  def gripper_to_mm(value_gripper, gripper_socket):
      closed_norm = get_closed_norm(gripper_socket)
      open_norm = get_open_norm(gripper_socket)
      closed_mm = get_closed_mm(gripper_socket)
      open_mm = get_open_mm(gripper_socket)

      value_norm = (value_gripper / 255) * 100

      slope = (closed_mm - open_mm) / (closed_norm - open_norm)
      value_mm = slope * (value_norm - closed_norm) + closed_mm

      if (value_mm > open_mm):
          value_mm_limited = open_mm
      elif (value_mm < closed_mm):
          value_mm_limited = closed_mm
      else:
          value_mm_limited = value_mm
      end

      return value_mm_limited
  end

  def mm_to_gripper(value_mm, gripper_socket):
      closed_norm = get_closed_norm(gripper_socket)
      open_norm = get_open_norm(gripper_socket)
      closed_mm = get_closed_mm(gripper_socket)
      open_mm = get_open_mm(gripper_socket)

      slope = (closed_norm - open_norm) / (closed_mm - open_mm)
      value_norm = (value_mm - closed_mm) * slope + closed_norm

      value_gripper = value_norm * 255 / 100

      if (value_gripper > 255):
          value_gripper_limited = 255
      elif (value_gripper < 0):
          value_gripper_limited = 0
      else:
          value_gripper_limited = round_value(value_gripper)
      end

      return value_gripper_limited
  end

  def round_value(value):
      value_mod = value % 1

      if(value_mod < 0.5):
          return floor(value)
      else:
          return ceil(value)
      end
  end

  def round_value_2_dec(value):
      value_x_100 = value * 100
      value_x_100_rounded = round_value(value_x_100)
      return value_x_100_rounded / 100
  end

  def clear_socket_buffer(gripper_socket="1", read_timeout = 0.1):
      rq_comm_clear_socket_buffer_enabled[rq_socket_to_index(gripper_socket)] = True
  end

  def rq_gripper_id_to_ascii(gripper_id):
      if(gripper_id == "1"):
          return 57
      elif(gripper_id == "2"):
          return 50
      elif(gripper_id == "3"):
          return 51
      elif(gripper_id == "4"):
          return 52
      end
  end

      def scale(value, rawRange, scaledRange):
          def computeSlope(inputRange, outputRange):
              outputRangeDelta = outputRange[1] - outputRange[0]
              inputRangeDelta = inputRange[1] - inputRange[0]

              if (inputRangeDelta == 0):
                  return 0
              else:
                  return outputRangeDelta / inputRangeDelta
              end
          end

          def computeIntercept(slope, inputRange, outputRange):
              return outputRange[0] - (slope * inputRange[0])
          end

          def clipScaledValue(outputScaledValue, outputRange):
              if (outputRange[0] < outputRange[1]):
                  return clipWhenLowerLimitIsLessThanHigher(outputScaledValue, outputRange)
              else:
                  return clipWhenLowerLimitIsGreaterThanHigherLimit(outputScaledValue, outputRange)
              end
          end

          def clipWhenLowerLimitIsGreaterThanHigherLimit(outputScaledValue, outputRange):
              if (outputScaledValue < outputRange[1]):
                  return outputRange[1]
              elif (outputScaledValue > outputRange[0]):
                  return outputRange[0]
              else:
                  return outputScaledValue
              end
          end

          def clipWhenLowerLimitIsLessThanHigher(outputScaledValue, outputRange):
              if (outputScaledValue < outputRange[0]):
                  return outputRange[0]
              elif (outputScaledValue > outputRange[1]):
                  return outputRange[1]
              else:
                  return outputScaledValue
              end
          end

          slope = computeSlope(rawRange, scaledRange)
          intercept = computeIntercept(slope, rawRange, scaledRange)
          scaledValue = slope * value + intercept
          return clipScaledValue(scaledValue, scaledRange)
      end

      def limit(value, range):
          return scale(value, range, range)
      end


  rq_init_comm_if_connected(9, "1")
  rq_init_comm_if_connected(2, "2")
  rq_init_comm_if_connected(3, "3")
  rq_init_comm_if_connected(4, "4")
  rq_print_connected_grippers()
  rq_gripper_communication_thread = run rq_gripper_communication()
  set_closed_norm(97.6470588235294, "1")
  set_open_norm(1.1764705882352942, "1")
  set_closed_mm(0.0, "1")
  set_open_mm(53.0, "1")
  set_closed_norm(100.0, "2")
  set_open_norm(0.0, "2")
  set_closed_mm(0.0, "2")
  set_open_mm(50.0, "2")
  set_closed_norm(100.0, "3")
  set_open_norm(0.0, "3")
  set_closed_mm(0.0, "3")
  set_open_mm(50.0, "3")
  set_closed_norm(100.0, "4")
  set_open_norm(0.0, "4")
  set_closed_mm(0.0, "4")
  set_open_mm(50.0, "4")
  rq_current_limit_enabled = False
  while(not rq_gripper_communication_thread_started):
      sleep(0.008)
  end
  # end: URCap Installation Node
  step_count_af30497c_f8d6_4abb_9ab3_badfcb3aff49 = 0.0
  thread Step_Counter_Thread_6e0f90e9_d7f0_45c2_bba1_3f0a34dad08c():
    while (True):
      step_count_af30497c_f8d6_4abb_9ab3_badfcb3aff49 = step_count_af30497c_f8d6_4abb_9ab3_badfcb3aff49 + 1.0
      sync()
    end
  end
  run Step_Counter_Thread_6e0f90e9_d7f0_45c2_bba1_3f0a34dad08c()
  global AMR_Position=struct(position_identifier=0, x1=0, x2=0, y1=0, y2=0, theta1=0, theta2=0)
  global CAM_Pose=p[0,0,0,0,0,0]
  global CAM_Relation=""
  global CMD_Abort=  False
  global CMD_Clear=  False
  global CMD_Reset=  False
  global CMD_Start=  False
  global CMD_Suspend=  False
  global CMD_Unhold=  False
  global CMD_Unsuspend=  False
  global CNT_Rack_Output=0
  global FNC_Freedrive=  False
  global PRC_TubCounter=0
  global STP=0
  global easyPickCount_4=0
  global easyPickCount_7=0
  global easyPickNoObj_4=0
  global easyPickNoObj_7=0
  global easyPickParts_4=0
  global easyPickParts_7=0
  global TMR_Barcode=0
  global Container_mid_1_p=p[-.379239199143, -.127191311915, .299999999998, .000000000046, -.000000000021, -1.247199999994]
  global Container_mid_1_q=[-2.477408934449926, -1.2969853503591224, -1.875639182904262, -1.539621866126728, 1.5731943360401213, -2.8009955944022717]
  global trigger_otw_p=p[-.364831738276, -.163967193938, .343299997821, .000000000046, -.000000000020, -1.148401333327]
  global trigger_otw_q=[-2.378283213085033, -1.2994862387706814, -1.7634300687554951, -1.6493302004167063, 1.573123683454141, -2.8011223671816943]
  global Waypoint_54_p=p[.008800512419, -.547926542621, .402696567415, -.589884378425, -.007228654778, -.061268144704]
  global Waypoint_54_q=[-1.2044575850116175, -1.3416667741588135, -1.8272563219070435, -0.9884541195682068, 1.3621035814285278, -2.7712565104113978]
  global Waypoint_77_p=p[-.178371829612, -.433927395311, .368082383916, -.086593488055, .704679941724, -.007869906074]
  global Waypoint_77_q=[-1.265390698109762, -1.3355963987163086, -1.7944865226745605, -1.7402602634825648, 0.8780410885810852, -2.7713127771960657]
  global Waypoint_83_p=p[.008800512419, -.547926542621, .402696567415, -.589884378425, -.007228654778, -.061268144704]
  global Waypoint_83_q=[-1.2044575850116175, -1.3416667741588135, -1.8272563219070435, -0.9884541195682068, 1.3621035814285278, -2.7712565104113978]
  global Waypoint_84_p=p[-.178371829612, -.433927395311, .368082383916, -.086593488055, .704679941724, -.007869906074]
  global Waypoint_84_q=[-1.265390698109762, -1.3355963987163086, -1.7944865226745605, -1.7402602634825648, 0.8780410885810852, -2.7713127771960657]
  global Vial_above_1_p=p[.017105793010, -.652093028359, .184920586844, .000000000272, .000000000270, 1.564063451276]
  global Vial_above_1_q=[-1.3375440709712851, -1.9618096977868804, -1.4665759083780685, -1.2837941559171444, 1.5732503672317195, -4.47276330421513]
  global Vial_pick_poi_1_p=p[.017105792852, -.648922724010, .093307568731, .000000000271, .000000000270, 1.564063451276]
  global Vial_pick_poi_1_q=[-1.3366329456391917, -2.0375277831965413, -1.6071432798879028, -1.0675084332049813, 1.57309887265915, -4.471135348858068]
  global Waypoint_86_p=p[.019227646885, -.648669633640, .184920586950, .000000000000, .000000000000, .024063451426]
  global Waypoint_86_q=[-1.3331129109407733, -1.9540750545686123, -1.4775914902901128, -1.280581784992414, 1.5733500744865856, -2.928303704452631]
  global Waypoint_87_p=p[-.032361834699, -.348336136197, .391475576335, -.000008499254, .000014589902, -.004651426820]
  global Waypoint_87_q=[-1.2709335019096129, -1.1914598663441005, -1.708995335060501, -1.8117888533498316, 1.5729683532263925, -2.8379347397710237]
  global Vial_3FG_plac_1_p=p[-.031858676359, -.349402499566, .145301120695, .000000000000, .000000000000, .000000000000]
  global Vial_3FG_plac_1_q=[-1.2723975525801707, -1.252376585823825, -2.3128114007049496, -1.1470592278900167, 1.5730548099411423, -2.8414815174610535]
  global Waypoint_88_p=p[-.032361834699, -.348336136197, .391475576335, -.000008499254, .000014589902, -.004651426820]
  global Waypoint_88_q=[-1.2709335019096129, -1.1914598663441005, -1.708995335060501, -1.8117888533498316, 1.5729683532263925, -2.8379347397710237]
  global cap_dump_1_p=p[-.139168676487, -.420163541420, .146096395183, .000000000000, .000000000000, .000000000000]
  global cap_dump_1_q=[-1.584588644510994, -1.5093464179777323, -2.1118449369620347, -1.091059703602438, 1.5728943834877336, -3.154014906686923]
  global Waypoint_89_p=p[-.032361834699, -.348336136197, .391475576335, -.000008499254, .000014589902, -.004651426820]
  global Waypoint_89_q=[-1.2709335019096129, -1.1914598663441005, -1.708995335060501, -1.8117888533498316, 1.5729683532263925, -2.8379347397710237]
  global Vial_3FG_plac_2_p=p[-.031858676359, -.349402499566, .145301120695, .000000000000, .000000000000, .000000000000]
  global Vial_3FG_plac_2_q=[-1.2723975525801707, -1.252376585823825, -2.3128114007049496, -1.1470592278900167, 1.5730548099411423, -2.8414815174610535]
  global Waypoint_90_p=p[-.032361834699, -.348336136197, .391475576335, -.000008499254, .000014589902, -.004651426820]
  global Waypoint_90_q=[-1.2709335019096129, -1.1914598663441005, -1.708995335060501, -1.8117888533498316, 1.5729683532263925, -2.8379347397710237]
  global cap_dump_2_p=p[-.139168676487, -.420163541420, .146096395183, .000000000000, .000000000000, .000000000000]
  global cap_dump_2_q=[-1.584588644510994, -1.5093464179777323, -2.1118449369620347, -1.091059703602438, 1.5728943834877336, -3.154014906686923]
  global Waypoint_91_p=p[-.032361834699, -.348336136197, .391475576335, -.000008499254, .000014589902, -.004651426820]
  global Waypoint_91_q=[-1.2709335019096129, -1.1914598663441005, -1.708995335060501, -1.8117888533498316, 1.5729683532263925, -2.8379347397710237]
  global Vial_liq_abov_1_p=p[-.025303660977, -.338758622354, .426628485936, -1.315858642253, .800043520260, -.928295855026]
  global Vial_liq_abov_1_q=[-0.3789628187762659, -1.5149522957256814, -2.263045310974121, 0.7870649534412841, -0.750984017048971, -3.2237566153155726]
  global Vial_liq_pick_3_p=p[-.002660428945, -.335984893034, .159389832934, -1.150456778400, .673175527684, -1.010612657503]
  global Vial_liq_pick_3_q=[-0.3660772482501429, -1.4503649038127442, -2.4056053161621094, -1.994692941705221, 0.8039668202400208, -0.2508929411517542]
  global Vial_liq_pick_4_p=p[-.041402486291, -.356791603314, .125395323246, -1.143483969075, .651070210027, -.878721885453]
  global Vial_liq_pick_4_q=[-0.4426233705502476, -1.437252121513727, -2.551930962114307, -1.776528229806984, 0.6562026234073748, -0.43018811960029524]
  global Vial_liq_abov_2_p=p[-.025303660977, -.338758622354, .426628485936, -1.315858642253, .800043520260, -.928295855026]
  global Vial_liq_abov_2_q=[-0.3789628187762659, -1.5149522957256814, -2.263045310974121, 0.7870649534412841, -0.750984017048971, -3.2237566153155726]
  global Liquid_midway_1_p=p[.057575295009, -.583081747994, .306414980749, -1.351675548728, .120935756539, -.096908606303]
  global Liquid_midway_1_q=[-0.895174805318014, -1.7035466633238734, -2.380953073501587, 0.631549521083496, 0.7706599235534668, -2.9455552736865442]
  global shake_3_p=p[.057574880217, -.583085370269, .306422893466, -1.360996190983, -.155555042453, -.438136255921]
  global shake_3_q=[-0.8951800505267542, -1.7035466633238734, -2.380937099456787, 0.6315542894550782, 0.7706599235534669, -2.5394540616517496]
  global shake_4_p=p[.057581636113, -.583090570002, .306439684073, -1.308767904323, .368530312677, .214926493520]
  global shake_4_q=[-0.8951714674579065, -1.7035395107665003, -2.380906343460083, 0.6315504747578125, 0.7706480026245118, -3.3161255787892268]
  global drop_above_3_p=p[.268235025993, -.467784390499, .226219872376, -1.027832627524, -.430841408251, 1.004603115937]
  global drop_above_3_q=[-0.935645882283346, -1.6663371525206507, -2.4252893924713135, 0.41966931402172847, 1.8470635414123535, -3.4600217978106897]
  global drop_above_4_p=p[.219042229014, -.470775657081, .133754190740, -.313004595901, -.344395319364, 1.500564994056]
  global drop_above_4_q=[-1.0601594887284795, -1.70046459045642, -2.0799996233759863, -0.7243227230676759, 1.9429634314685202, -4.115129153870795]
  global liq_tran_3_p=p[.213067510942, -.469567035397, .100231043184, .251862243732, .217902579404, 1.592812335393]
  global liq_tran_3_q=[-0.7789645168037476, -1.822364827406652, -1.8643518410805573, -1.252158963840138, 1.3768134449520435, -3.9328333233290254]
  global drop_above_5_p=p[.219042229014, -.470775657081, .133754190740, -.313004595901, -.344395319364, 1.500564994056]
  global drop_above_5_q=[-1.0601594887284795, -1.70046459045642, -2.0799996233759863, -0.7243227230676759, 1.9429634314685202, -4.115129153870795]
  global Waypoint_92_p=p[.187119460405, -.493959476151, .133754190608, -.313004596540, -.344395317757, 1.500564993991]
  global Waypoint_92_q=[-1.1418328121400876, -1.7310553375189475, -2.033634768766424, -0.772026910513711, 1.958578934631971, -4.201588449364511]
  global liq_tran_4_p=p[.195957706507, -.493022614126, .100231042689, .160718757180, .109807038912, 1.525321508623]
  global liq_tran_4_q=[-0.881740380645474, -1.8244526267589851, -1.865100964490387, -1.1608866323693583, 1.4631433601076713, -3.973915130363038]
  global drop_above_6_p=p[.219042229014, -.470775657081, .133754190740, -.313004595901, -.344395319364, 1.500564994056]
  global drop_above_6_q=[-1.0601594887284795, -1.70046459045642, -2.0799996233759863, -0.7243227230676759, 1.9429634314685202, -4.115129153870795]
  global drop_above_7_p=p[.268235025993, -.467784390499, .226219872376, -1.027832627524, -.430841408251, 1.004603115937]
  global drop_above_7_q=[-0.935645882283346, -1.6663371525206507, -2.4252893924713135, 0.41966931402172847, 1.8470635414123535, -3.4600217978106897]
  global Liquid_midway_2_p=p[.057575295009, -.583081747994, .306414980749, -1.351675548728, .120935756539, -.096908606303]
  global Liquid_midway_2_q=[-0.895174805318014, -1.7035466633238734, -2.380953073501587, 0.631549521083496, 0.7706599235534668, -2.9455552736865442]
  global Vial_drop_abo_1_p=p[.000324902251, -.648569523142, .221894115667, -.873462921366, 1.165852672573, -1.482720593185]
  global Vial_drop_abo_1_q=[-1.0576906334721352, -2.393016994184633, -0.9236232851859159, -2.5729213042279273, 0.7903331288549689, -0.33286325848155585]
  global Vial_liq_drop_1_p=p[.001020867953, -.647659915585, .092915870838, -.834762611599, 1.081942994823, -1.540647900176]
  global Vial_liq_drop_1_q=[-1.0631954168193474, -2.4447642951220825, -1.128811017825127, -2.1983115491972294, 0.8130148661460634, -0.38984988696911316]
  global Vial_drop_abo_2_p=p[.000324902251, -.648569523142, .221894115667, -.873462921366, 1.165852672573, -1.482720593185]
  global Vial_drop_abo_2_q=[-1.0576906334721352, -2.393016994184633, -0.9236232851859159, -2.5729213042279273, 0.7903331288549689, -0.33286325848155585]
  global Spatula_otw_p=p[-.038472058237, -.263141484147, .425351216717, -.000441582511, -.000128175490, 3.034387645854]
  global Spatula_otw_q=[-1.1888947506684495, -1.0083288774886814, -1.7052227056065874, -1.9984805067363443, 1.5730180972985317, 0.48793409320312264]
  global pick_spat_L_abv_p=p[.239059466375, -.067212518441, .280720723617, .000017217488, -.000484427718, 3.106837214660]
  global pick_spat_L_abv_q=[0.292765616142962, -0.8565557553273315, -2.140199892763044, -1.715349495646084, 1.573623142106424, 1.8984976776985687]
  global spat_L_pick_p=p[.242468789885, -.067301915011, .193171208067, .000017217488, -.000484427718, 3.106837214657]
  global spat_L_pick_q=[0.2867414378807389, -0.8600077002089179, -2.3629148016312627, -1.4891831672860159, 1.5737695566221115, 1.8933890858591198]
  global spat_L_lift_p=p[.245402002494, -.067432373551, .289049296496, .000017217490, -.000484427724, 3.106837214657]
  global spat_L_lift_q=[0.2834351187564135, -0.8798320076811592, -2.1119436738532986, -1.7203314352121302, 1.573588313403067, 1.8891054681654005]
  global spat_L_side_p=p[.247133573905, -.017633681797, .289062935631, .000017217490, -.000484427724, 3.106837214657]
  global spat_L_side_q=[0.49719173575848863, -0.8582398211168538, -2.1182130454788215, -1.735610316654931, 1.5735817737572706, 2.1028402698705397]
  global spat_L_up_p=p[.247135508752, -.017665230822, .397130746165, .000017217490, -.000484427724, 3.106837214657]
  global spat_L_up_q=[0.49854946074076967, -0.9346239623559676, -1.808280269374471, -1.969158816463132, 1.5731020084036995, 2.1031742024348157]
  global spat_M_up_p=p[.244670000000, -.112000000000, .420343789747, .000026293990, -.000477463070, 3.067686800857]
  global spat_M_up_q=[0.09097498152209688, -1.0114245603211778, -1.718034632879454, -1.9826932847219538, 1.5730130135866505, 1.734554438783734]
  global spat_M_pick_p=p[.244673518506, -.111985070134, .192299022723, .000043885692, -.000001622442, 3.067686841404]
  global spat_M_pick_q=[0.08868170265231701, -0.9271392933223233, -2.343826449241451, -1.441236864368305, 1.5733923850045939, 1.7345552462242537]
  global spat_S_Up_7_p=p[.243228810603, -.161948321982, .423281604617, .000026293955, -.000477463064, 3.067686800854]
  global spat_S_Up_7_q=[-0.11182322368059516, -1.0716267311491734, -1.6854498186860427, -1.955120134033855, 1.5730106579635699, 1.5317349120701778]
  global spat_S_Pick_4_p=p[.245377020686, -.158668022535, .192285730279, .000026293985, -.000477463062, 3.067686800840]
  global spat_S_Pick_4_q=[-0.10087203759495189, -1.011188488703386, -2.311978084495874, -1.3890267520590838, 1.5735990551056096, 1.5450562970948172]
  global spat_S_Up_8_p=p[.252087445596, -.159242094834, .423281604617, .000026293954, -.000477463070, 3.067686800855]
  global spat_S_Up_8_q=[-0.09804692328730358, -1.0862987822056382, -1.6788706463996483, -1.9470242450550348, 1.5730147401359813, 1.5455107082823842]
  global spat_flatM_up_p=p[.241028517126, -.208127630016, .404671074680, .000026293951, -.000477463078, 3.067686800891]
  global spat_flatM_up_q=[-0.27878462628263456, -1.1217510366315881, -1.7121530048618725, -1.8783279876432832, 1.5731053960668042, 1.3649536117980254]
  global spat_flatM_pick_p=p[.241028983327, -.208057297586, .192270533170, .000026293950, -.000477463079, 3.067686800885]
  global spat_flatM_pick_q=[-0.2805687960562633, -1.1003763929487214, -2.271431297337675, -1.3404236887924883, 1.5734924238720627, 1.3653813047742556]
  global spat_flatS_up_p=p[.237651953780, -.253943828614, .403961222825, .000026293950, -.000477463092, 3.067686800841]
  global spat_flatS_up_q=[-0.42363550926974103, -1.1939944599502539, -1.6745915127240307, -1.843675057902054, 1.5731001874678698, 1.220082820532415]
  global spat_flatS_pick_p=p[.241325662334, -.251726327528, .192256842740, .000026293947, -.000477463087, 3.067686800841]
  global spat_flatS_pick_q=[-0.4144907797170738, -1.1967447109013012, -2.21926362252748, -1.2962499335425761, 1.5733885098427622, 1.2314402238866728]
  global spat_S_pick_p=p[.241585614619, -.158882677087, .191636172448, .000019478956, -.000483249177, 3.097147973434]
  global spat_S_pick_q=[-0.10320942227973173, -1.0007485193115802, -2.317947069452162, -1.3934956127505886, 1.5736112980229278, 1.5132597021160705]
  global spat_S_up_p=p[.248189103503, -.159371150053, .417088864416, .000026293966, -.000477463070, 3.067686800840]
  global spat_S_up_q=[-0.10007737460061872, -1.0730270029702904, -1.7018049146034766, -1.9373622285571734, 1.573045444550866, 1.5435422173047084]
  global Waypoint_7_p=p[-.472820924474, .292439826233, .207418370237, -.137787250486, 2.177332259632, -2.152029714756]
  global Waypoint_7_q=[-2.911134078210732, -1.90240864358569, -1.968768330510411, -2.500365101593811, 0.11427687110891149, 0.0958980389250167]
  global Waypoint_8_p=p[-.357612884176, -.251084817998, .212379799667, -.858181193174, 1.714832512191, -1.687547565568]
  global Waypoint_8_q=[-1.620834863369681, -1.8936194567376496, -1.9821394403832038, -2.4599791457905273, 0.6296693672615152, 0.07625365420707819]
  global Decapp_above_3_p=p[-.013480295948, -.359153355979, .266194408367, -.879653555922, 1.646336924805, -1.709111068605]
  global Decapp_above_3_q=[-0.9632157249872035, -2.0163405763031657, -1.5968194594157152, -2.6579215719847085, 1.251243398585566, 0.047906446502667066]
  global Decapp_place_3_p=p[-.013480295890, -.359153356055, .160907502384, -.879653554902, 1.646336919740, -1.709111066456]
  global Decapp_place_3_q=[-0.9633402410919709, -2.1541179572356635, -1.6937729380888573, -2.4232786481058053, 1.2517342187662468, 0.04818402956922263]
  global Decapp_above_4_p=p[-.013480295948, -.359153355979, .266194408367, -.879653555922, 1.646336924805, -1.709111068605]
  global Decapp_above_4_q=[-0.9632157249872035, -2.0163405763031657, -1.5968194594157152, -2.6579215719847085, 1.251243398585566, 0.047906446502667066]
  global Waypoint_78_p=p[-.051450028091, -.519555688329, .365718563414, -1.287302938145, 1.077637394477, -1.218524965834]
  global Waypoint_78_q=[-0.9214276262416012, -1.8899696965062578, -1.4939326452510562, -2.840015661555725, 0.5585157189668353, 0.033997638875617575]
  global Waypoint_10_p=p[-.466751210260, .252836712095, .259921246286, 1.042686976164, .439333316918, -1.691967798809]
  global Waypoint_10_q=[-3.022216346250036, -1.8383597675135919, -1.566977059184386, -2.046864464116096, 0.8487467526238, -2.4392912369481916]
  global Waypoint_9_p=p[-.538777454962, .370695704977, .175030018143, -.317104215445, 2.082346543003, -2.037631421082]
  global Waypoint_9_q=[-3.1158871966457857, -1.998548595120492, -1.941797010061462, -2.2703530575838844, -0.27573365931009164, -0.06926782177267654]
  global Powder_wayp1_p=p[-.472820924474, .292439826233, .207418370237, -.137787250486, 2.177332259632, -2.152029714756]
  global Powder_wayp1_q=[-2.911134078210732, -1.90240864358569, -1.968768330510411, -2.500365101593811, 0.11427687110891149, 0.0958980389250167]
  global Waypoint_2_p=p[-.357612884176, -.251084817998, .212379799667, -.858181193174, 1.714832512191, -1.687547565568]
  global Waypoint_2_q=[-1.620834863369681, -1.8936194567376496, -1.9821394403832038, -2.4599791457905273, 0.6296693672615152, 0.07625365420707819]
  global Postions_otw_p=p[-.010896578244, -.533368729951, .288851175116, -1.233738470894, 1.195331112012, -1.207314088469]
  global Postions_otw_q=[-0.898791023514228, -2.078490033037677, -1.4499891355755317, -2.7624416226992476, 0.6570218891920963, 0.02136606178275929]
  global cont_A_otw_p=p[.070238108556, -.655257851554, .184611566008, -1.090601381517, 1.404822685081, -1.413645380264]
  global cont_A_otw_q=[-0.990969136335913, -2.7123780097559784, -0.5772671651193146, -3.0005537851220403, 0.84719335943793, 0.020652463706785973]
  global cont_B_otw_p=p[.255895686750, -.501120003087, .157855243207, -1.209177187561, 1.209243088037, -1.209202949417]
  global cont_B_otw_q=[-0.5819602570351563, -2.5181180937953833, -1.0264696604583161, -2.7360726814058687, 0.9880932038785559, -0.004134033524621827]
  global cont_B_safe_p=p[.242897168204, -.501733713795, .237745474779, -1.209212324107, 1.209144328638, -1.209309913894]
  global cont_B_safe_q=[-0.5929699566143585, -2.4210115429142114, -0.9949203644592259, -2.8646436479104267, 0.976678899749076, -0.004020526358775811]
  global cont_C_otw_p=p[.319495487998, -.362719410364, .163846736977, -1.233784872294, 1.195277203291, -1.207325031551]
  global cont_C_otw_q=[-0.3611889651645974, -2.404603865546651, -1.2341573845076566, -2.650535279811077, 1.1944844573128257, 0.01638086594640864]
  global Waypoint_1_p=p[-.352029261722, -.424157832422, .472326578019, -.000004407962, .000020663369, -1.529709227737]
  global Waypoint_1_q=[-2.017015745614491, -1.7423968528991196, -1.0053357238485425, -1.9644715035904907, 1.5727249689896, -2.060727852912713]
  global Waypoint_5_p=p[.219993437017, -.447144142811, .462350040687, .000006087494, .000031090075, .000022232405]
  global Waypoint_5_q=[-0.8406239476037944, -1.5982534362206806, -1.1934200873248484, -1.9205794898315975, 1.5727336676986443, -2.4135960466995314]
  global place_2_home_p=p[-.352029261717, -.424157832411, .329197314759, -.000004407962, .000020663369, -1.529709227737]
  global place_2_home_q=[-2.017880982348384, -1.6708952803108668, -1.462293789471877, -1.5790150659586653, 1.5732060241635952, -2.059940179665328]
  global Waypoint_12_p=p[-.812560029877, -.415067232840, .258518340146, -1.257569567036, 1.159670338548, -1.145019586130]
  global Waypoint_12_q=[-2.3224548809497123, -2.3211405271930765, -1.1304722687551445, -2.8155296475017018, -0.8321758827962036, -0.007205995478960503]
  global Waypoint_18_p=p[-.813643087636, -.416224939441, .099970000000, -1.257570310935, 1.159676546330, -1.145010619029]
  global Waypoint_18_q=[-2.322494764677227, -2.501268559301314, -1.239250885783676, -2.5265468980680197, -0.831327849164623, -0.00732105677136996]
  global Waypoint_19_p=p[-.812560029269, -.415067232191, .079455005744, -1.257569567033, 1.159670338546, -1.145019586137]
  global Waypoint_19_q=[-2.3224951834453367, -2.5274729453886575, -1.2489176533831348, -2.4906644180980346, -0.8312252662037514, -0.007338111970053518]
  def calculate_point_to_move_towards(feature, direction, position_distance):
    local posDir=[direction[0], direction[1], direction[2]]
    if (norm(posDir) < 1e-6):
      return get_target_waypoint()
    end
    local direction_vector_normalized=normalize(posDir)
    local displacement_pose=p[direction_vector_normalized[0] * position_distance,direction_vector_normalized[1] * position_distance,direction_vector_normalized[2] * position_distance,0,0,0]
    local wanted_displacement_in_base_frame=pose_sub(pose_trans(feature, displacement_pose), feature)
    return pose_add(get_target_waypoint(), wanted_displacement_in_base_frame)
  end
  global TMR_Barcode_is_counting=False
  thread Timer_Thread():
    while (True):
      if (TMR_Barcode_is_counting):
        TMR_Barcode = TMR_Barcode + get_steptime()
      end
      sync()
    end
  end
  run Timer_Thread()
  def Sub_Vision_V18():
    $ 892 "Sub_Vision_V18" "noBreak"
    $ 893 "PreSettings"
    $ 894 "CAM_LM_Detected≔ False "
    global CAM_LM_Detected=  False
    $ 895 "CAM_Captures≔0"
    global CAM_Captures=0
    $ 896 "CAM_Pose≔p[0,0,0,0,0,0]"
    global CAM_Pose=p[0,0,0,0,0,0]
    $ 897 "CAM_LM_Refinmnt≔ False "
    global CAM_LM_Refinmnt=  False
    $ 898 "CAM_LM_Refined≔ False "
    global CAM_LM_Refined=  False
    $ 899 "CAM_LM_Deviatn≔p[0,0,0,0,0,0]"
    global CAM_LM_Deviatn=p[0,0,0,0,0,0]
    $ 900 "CAM_LM_ID≔0"
    global CAM_LM_ID=0
    $ 901 "CAM_Done≔ False "
    global CAM_Done=  False
    $ 902 "CAM_CNT_Obj≔0"
    global CAM_CNT_Obj=0
    $ 903 "CAM_Result = []"
    CAM_Result = []
    $ 904 "OBJ_Detected≔ False "
    global OBJ_Detected=  False
    $ 905 "FRM_Reference≔p[0,0,0,0,0,0]"
    global FRM_Reference=p[0,0,0,0,0,0]
    $ 906 "'=========='"
    # '=========='
    $ 907 "Switch Action"
    switch_1 = Action
    $ 908 "Case 13"
    if (13 == switch_1):
    elif (15 == switch_1):
      $ 1026 "Case 15"
    elif (131 == switch_1):
      $ 1072 "Case 131"
      $ 1073 "Read (SensoPart)"
      $ 1074 "Action_Info≔'search for landmark'"
      global Action_Info="search for landmark"
      $ 1075 "CAM_LM≔CAM_LMs[4]"
      global CAM_LM=CAM_LMs[4]
      $ 1076 "CAM_Relation≔CAM_LM.capture_relation"
      global CAM_Relation=CAM_LM.capture_relation
      $ 1077 "go to capture pose"
      $ 1080 "If ITM_ID≟1 and JIG≟7"
      if (ITM_ID == 1  and  JIG == 7):
        $ 1081 "PSE_T≔uLM_Cap_SSRack"
        global PSE_T=uLM_Cap_SSRack
      else:
        $ 1082 "ElseIf ITM_ID≟5 and JIG≟7"
        if (ITM_ID == 5  and  JIG == 7):
          $ 1083 "PSE_T≔FRM_Cap_SSRack"
          global PSE_T=FRM_Cap_SSRack
        else:
          $ 1086 "ElseIf ITM_ID≟1 and JIG≟15"
          if (ITM_ID == 1 and JIG == 15):
            $ 1087 "MoveJ"
            $ 1088 "Container_mid_1" "breakAfter"
            movej(get_inverse_kin(Container_mid_1_p, qnear=Container_mid_1_q), a=1.3962634015954636, v=1.0471975511965976, r=0.05)
            $ 1090 "PSE_T≔FRM_Container_const"
            global PSE_T=p[-0.5003348223692186,0.35061804815168285,0.41579001388808423,-5.092943187272062E-5,1.0145185065363121E-4,-2.764319258713288]
          else:
            $ 1091 "ElseIf ITM_ID≟1 and JIG≟21"
            if (ITM_ID == 1 and JIG == 21):
              $ 1093 "PSE_T≔FRM_PoTS_const"
              global PSE_T=p[-0.5403054403210852,-0.10910773999775857,0.4828,3.058497512721046E-6,2.3454853329357316E-5,-2.208510541952706]
            else:
              $ 1094 "ElseIf ITM_ID≟1 and JIG≟22"
              if (ITM_ID == 1 and JIG == 22):
                $ 1096 "MoveJ"
                $ 1097 "FRM_PoTS" "breakAfter"
                movej(FRM_PoTS, a=1.3962634015954636, v=1.0471975511965976, r=0.05)
                $ 1098 "PSE_T≔FRM_SWAB_const"
                global PSE_T=p[-0.5425658438438228,0.050215382883637555,0.4828117991467299,1.2014498510989115E-5,1.8611655946156755E-5,-2.2084947047695405]
              else:
                $ 1099 "ElseIf ITM_ID≟1 and JIG≟17"
                if (ITM_ID == 1 and JIG == 17):
                  $ 1100 "MoveJ"
                  $ 1101 "zero_scale()"
                  zero_scale()
                  $ 1102 "trigger_otw" "breakAfter"
                  movej(get_inverse_kin(trigger_otw_p, qnear=trigger_otw_q), a=1.3962634015954636, v=1.0471975511965976, r=0.05)
                  $ 1106 "PSE_T≔FRM_weigh_scale_const"
                  global PSE_T=p[-0.3804866881697204,0.025744252835212,0.4723487455232425,-1.0445769542396123E-4,-1.924788411074358E-5,-2.1691978730572363]
                end
              end
            end
          end
        end
      end
      $ 1107 "do_transition(PSE_T, keep_rxry=False)"
      do_transition(PSE_T, keep_rxry=False)
      $ 1108 "Set"
      set_tcp(p[0.0,0.0,0.161,3.1415,0.0,0.0])
      $ 1109 "MoveJ"
      $ 1110 "PSE_T" "breakAfter"
      movej(PSE_T, a=1.3962634015954636, v=1.7453292519943295)
      $ 1111 "CAM_Pose≔get_actual_tcp_pose()"
      global CAM_Pose= get_actual_tcp_pose ()
      $ 1112 "Loop  not CAM_Done and  not ERROR.FLAG and  not CMD_Stop"
      while (  not  CAM_Done  and    not  ERROR.FLAG  and    not  CMD_Stop):
        $ 1113 "adjust capture pose"
        $ 1114 "If CAM_LM_Detected and CAM_LM_Refinmnt"
        if (CAM_LM_Detected  and  CAM_LM_Refinmnt):
          $ 1115 "PSE_T≔p[0,0,0.300,0,0,0]"
          global PSE_T=p[0,0,0.300,0,0,0]
          $ 1116 "CAM_Pose≔PSE_T"
          global CAM_Pose=PSE_T
          $ 1117 "If  not is_reachable(FRM_Reference,[PSE_T])"
          if (  not  is_reachable(FRM_Reference,[PSE_T])):
            $ 1118 "Error"
            $ 1119 "set_error(ERROR_POSE_NOT_REACHABLE)"
            set_error(ERROR_POSE_NOT_REACHABLE)
          end
          $ 1120 "If  not ERROR.FLAG"
          if (  not  ERROR.FLAG):
            $ 1121 "MoveJ"
            $ 1122 "PSE_T" "breakAfter"
            set_tcp(p[0.0,0.0,0.161,0.0,0.0,0.0])
            movej(pose_trans(FRM_Reference, PSE_T), a=0.8726646259971648, v=1.3962634015954636)
            $ 1123 "CAM_LM_Refined≔ True "
            global CAM_LM_Refined=  True
          end
        else:
          $ 1124 "ElseIf  not CAM_LM_Detected and CAM_Captures>0"
          if (  not  CAM_LM_Detected  and  CAM_Captures>0):
            $ 1125 "MoveL"
            $ 1126 "If FRM_Reference≟p[0,0,0,0,0,0]"
            if (FRM_Reference == p[0,0,0,0,0,0]):
              $ 1127 "PSE_T≔get_random_pose(pose_ref=CAM_Pose, mode='cubic', range_max=[0.150,0.150,0.015])"
              global PSE_T=get_random_pose(pose_ref=CAM_Pose, mode="cubic", range_max=[0.150,0.150,0.015])
            else:
              $ 1132 "Else" "noBreak"
              $ 1133 "PSE_T≔get_random_pose(pose_ref=CAM_Pose, mode='rotation', range_max=[10,10,0])"
              global PSE_T=get_random_pose(pose_ref=CAM_Pose, mode="rotation", range_max=[10,10,0])
              $ 1134 "CAM_LM_Refined≔ True "
              global CAM_LM_Refined=  True
            end
            $ 1135 "If get_inverse_kin_has_solution(pose_trans(FRM_Reference, PSE_T))"
            if (get_inverse_kin_has_solution( pose_trans (FRM_Reference, PSE_T))):
              $ 1136 "Comment"
              # Comment
              $ 1137 "PSE_T" "breakAfter"
              set_tcp(p[0.0,0.0,0.161,3.1415,0.0,0.0])
              movel(pose_trans(FRM_Reference, PSE_T), a=0.03, v=0.05)
            else:
              $ 1138 "Else" "noBreak"
              $ 1139 "'If random pose is out of reach, set the initial cam pose'"
              # 'If random pose is out of reach, set the initial cam pose'
              $ 1140 "PSE_T≔CAM_Pose"
              global PSE_T=CAM_Pose
            end
          end
        end
        $ 1141 "Wait: 2.0"
        sleep(2.0)
        $ 1142 "trigger"
        $ 1143 "If ITM_ID≟1 and JIG≟7"
        if (ITM_ID == 1  and  JIG == 7):
          # begin: URCap Program Node
          #   Source: SensoPart VISOR Robotic, 2.0.6, SensoPart Industriesensorik GmbH
          #   Type: VISOR Trigger
          $ 1144 "# 1 VISOR Trigger"
          visor_changeJob(1, "Landmark_INVITE_2", 6000)
          visor_trigger(1, 6000, "arm")
          # end: URCap Program Node
        else:
          $ 1145 "ElseIf ITM_ID≟5 and JIG≟7"
          if (ITM_ID == 5  and  JIG == 7):
            # begin: URCap Program Node
            #   Source: SensoPart VISOR Robotic, 2.0.6, SensoPart Industriesensorik GmbH
            #   Type: VISOR Trigger
            $ 1146 "# 1 VISOR Trigger"
            visor_changeJob(1, "Landmark_INVITE_2", 6000)
            visor_trigger(1, 6000, "arm")
            # end: URCap Program Node
          else:
            $ 1147 "ElseIf ITM_ID≟13 and JIG≟7"
            if (ITM_ID == 13  and  JIG == 7):
              # begin: URCap Program Node
              #   Source: SensoPart VISOR Robotic, 2.0.6, SensoPart Industriesensorik GmbH
              #   Type: VISOR Trigger
              $ 1148 "# 1 VISOR Trigger"
              visor_changeJob(1, "Landmark_INVITE_2", 6000)
              visor_trigger(1, 6000, "arm")
              # end: URCap Program Node
            else:
              $ 1149 "ElseIf ITM_ID≟1 and JIG≟15"
              if (ITM_ID == 1 and JIG == 15):
                # begin: URCap Program Node
                #   Source: SensoPart VISOR Robotic, 2.0.6, SensoPart Industriesensorik GmbH
                #   Type: VISOR Trigger
                $ 1150 "# 1 VISOR Trigger"
                visor_changeJob(1, "Aztec_no_dot_pick", 6000)
                visor_trigger(1, 6000, "arm")
                # end: URCap Program Node
              else:
                $ 1151 "ElseIf ITM_ID≟1 and JIG≟21"
                if (ITM_ID == 1 and JIG == 21):
                  # begin: URCap Program Node
                  #   Source: SensoPart VISOR Robotic, 2.0.6, SensoPart Industriesensorik GmbH
                  #   Type: VISOR Trigger
                  $ 1152 "# 1 VISOR Trigger"
                  visor_changeJob(1, "PoTS", 6000)
                  visor_trigger(1, 6000, "arm")
                  # end: URCap Program Node
                else:
                  $ 1153 "ElseIf ITM_ID≟1 and JIG≟17"
                  if (ITM_ID == 1 and JIG == 17):
                    # begin: URCap Program Node
                    #   Source: SensoPart VISOR Robotic, 2.0.6, SensoPart Industriesensorik GmbH
                    #   Type: VISOR Trigger
                    $ 1154 "# 1 VISOR Trigger"
                    visor_changeJob(1, "Weigh_target", 6000)
                    visor_trigger(1, 6000, "arm")
                    # end: URCap Program Node
                  else:
                    $ 1155 "ElseIf ITM_ID≟1 and JIG≟22"
                    if (ITM_ID == 1 and JIG == 22):
                      # begin: URCap Program Node
                      #   Source: SensoPart VISOR Robotic, 2.0.6, SensoPart Industriesensorik GmbH
                      #   Type: VISOR Trigger
                      $ 1156 "# 1 VISOR Trigger"
                      visor_changeJob(1, "Swab_Marker", 6000)
                      visor_trigger(1, 6000, "arm")
                      # end: URCap Program Node
                    end
                  end
                end
              end
            end
          end
        end
        $ 1160 "TM_3D_Found≔visor_partsFound(1)"
        global TM_3D_Found= visor_partsFound (1)
        $ 1162 "If TM_3D_Found>0"
        if (TM_3D_Found>0):
          $ 1163 "CAM_LM_Detected≔ True "
          global CAM_LM_Detected=  True
          $ 1164 "CAM_Captures≔0"
          global CAM_Captures=0
        else:
          $ 1165 "Else" "noBreak"
          $ 1166 "CAM_LM_Detected≔ False "
          global CAM_LM_Detected=  False
          $ 1167 "CAM_Captures≔CAM_Captures+1"
          global CAM_Captures=CAM_Captures+1
        end
        $ 1172 "result"
        $ 1173 "If CAM_LM_Detected"
        if (CAM_LM_Detected):
          $ 1174 "If (CAM_LM_Refinmnt and CAM_LM_Refined) or  not CAM_LM_Refinmnt"
          if ((CAM_LM_Refinmnt  and  CAM_LM_Refined)  or    not  CAM_LM_Refinmnt):
            $ 1232 "If ITM_ID≟1 and JIG≟7"
            if (ITM_ID == 1  and  JIG == 7):
              $ 1233 "CAM_LM_SSRack≔visor_getPose3d(1, 0)"
              global CAM_LM_SSRack= visor_getPose3d (1, 0)
            else:
              $ 1234 "ElseIf ITM_ID≟5 and JIG≟7"
              if (ITM_ID == 5  and  JIG == 7):
                $ 1235 "CAM_LM_SSRack≔visor_getPose3d(1, 0)"
                global CAM_LM_SSRack= visor_getPose3d (1, 0)
              else:
                $ 1238 "ElseIf ITM_ID≟1 and JIG≟15"
                if (ITM_ID == 1 and JIG == 15):
                  $ 1239 "CAM_LM_cont≔visor_getPose3d(1, 0)"
                  global CAM_LM_cont= visor_getPose3d (1, 0)
                  $ 1240 "Trigger≔get_actual_tcp_pose()"
                  global Trigger= get_actual_tcp_pose ()
                else:
                  $ 1241 "ElseIf ITM_ID≟1 and JIG≟21"
                  if (ITM_ID == 1 and JIG == 21):
                    $ 1242 "CAM_LM_cont≔visor_getPose3d(1, 0)"
                    global CAM_LM_cont= visor_getPose3d (1, 0)
                    $ 1243 "Trigger≔get_actual_tcp_pose()"
                    global Trigger= get_actual_tcp_pose ()
                  else:
                    $ 1244 "ElseIf ITM_ID≟1 and JIG≟17"
                    if (ITM_ID == 1 and JIG == 17):
                      $ 1245 "CAM_LM_cont≔visor_getPose3d(1, 0)"
                      global CAM_LM_cont= visor_getPose3d (1, 0)
                      $ 1246 "Trigger≔get_actual_tcp_pose()"
                      global Trigger= get_actual_tcp_pose ()
                    else:
                      $ 1247 "ElseIf ITM_ID≟1 and JIG≟22"
                      if (ITM_ID == 1 and JIG == 22):
                        $ 1248 "CAM_LM_cont≔visor_getPose3d(1, 0)"
                        global CAM_LM_cont= visor_getPose3d (1, 0)
                        $ 1249 "Trigger≔get_actual_tcp_pose()"
                        global Trigger= get_actual_tcp_pose ()
                      end
                    end
                  end
                end
              end
            end
            $ 1250 "CAM_Done≔ True "
            global CAM_Done=  True
          end
        else:
          $ 1251 "ElseIf  not CAM_LM_Detected and CAM_Captures<CAM_PRM_Retries"
          if (  not  CAM_LM_Detected  and  CAM_Captures<CAM_PRM_Retries):
            $ 1252 "CAM_LM_Refined≔ False "
            global CAM_LM_Refined=  False
          else:
            $ 1253 "ElseIf CAM_Captures≥CAM_PRM_Retries"
            if (CAM_Captures >= CAM_PRM_Retries):
              $ 1254 "CAM_Done≔ True "
              global CAM_Done=  True
              $ 1255 "Error"
              $ 1256 "set_error(ERROR_NO_LANDMARK)"
              set_error(ERROR_NO_LANDMARK)
            end
          end
        end
      end
    elif (151 == switch_1):
      $ 1257 "Case 151"
      $ 1258 "Detect (SensoPart)"
      $ 1259 "go to capture pose"
      $ 1260 "FRM_Reference≔FRM_Cap_SSRack"
      global FRM_Reference=FRM_Cap_SSRack
      $ 1261 "PSE_T≔p[0,0,-0.00,0,0,0]"
      global PSE_T=p[0,0,-0.00,0,0,0]
      $ 1262 "do_transition(pose_trans(FRM_Reference, PSE_T), keep_rxry=False)"
      do_transition( pose_trans (FRM_Reference, PSE_T), keep_rxry=False)
      $ 1263 "JNT_Q≔get_actual_joint_positions()"
      global JNT_Q= get_actual_joint_positions ()
      $ 1264 "JNT_Q≔[JNT_Q[0], JNT_Q[1], JNT_Q[2], JNT_Q[3], JNT_Q[4], 0]"
      global JNT_Q=[JNT_Q[0], JNT_Q[1], JNT_Q[2], JNT_Q[3], JNT_Q[4], 0]
      $ 1265 "Set"
      set_tcp(p[0.0,0.0,0.161,3.1415,0.0,0.0])
      $ 1266 "movej(get_inverse_kin(pose_trans(FRM_Reference, PSE_T), qnear=JNT_Q))"
      movej(get_inverse_kin( pose_trans (FRM_Reference, PSE_T), qnear=JNT_Q))
      $ 1267 "CAM_Pose≔pose_trans(pose_inv(FRM_Reference), get_actual_tcp_pose())"
      global CAM_Pose= pose_trans ( pose_inv (FRM_Reference),  get_actual_tcp_pose ())
      $ 1268 "Loop  not CAM_Done and  not ERROR.FLAG and  not CMD_Stop"
      while (  not  CAM_Done  and    not  ERROR.FLAG  and    not  CMD_Stop):
        $ 1269 "If  not OBJ_Detected and CAM_Captures>0"
        if (  not  OBJ_Detected  and  CAM_Captures>0):
          $ 1270 "MoveL"
          $ 1271 "If FRM_Reference≟p[0,0,0,0,0,0]"
          if (FRM_Reference == p[0,0,0,0,0,0]):
            $ 1273 "PSE_T≔get_random_pose(pose_ref=CAM_Pose, mode='rotation', range_max=[15,15,0])"
            global PSE_T=get_random_pose(pose_ref=CAM_Pose, mode="rotation", range_max=[15,15,0])
          else:
            $ 1274 "Else" "noBreak"
            $ 1275 "PSE_T≔get_random_pose(pose_ref=CAM_Pose, mode='rotation', range_max=[10,10,0])"
            global PSE_T=get_random_pose(pose_ref=CAM_Pose, mode="rotation", range_max=[10,10,0])
          end
          $ 1276 "If get_inverse_kin_has_solution(pose_trans(FRM_Reference, PSE_T))"
          if (get_inverse_kin_has_solution( pose_trans (FRM_Reference, PSE_T))):
            $ 1277 "PSE_T" "breakAfter"
            set_tcp(p[0.0,0.0,0.161,3.1415,0.0,0.0])
            movel(pose_trans(FRM_Reference, PSE_T), a=0.03, v=0.05)
          else:
            $ 1278 "Else" "noBreak"
            $ 1279 "'If random pose is out of reach, set the initial cam pose'"
            # 'If random pose is out of reach, set the initial cam pose'
            $ 1280 "PSE_T≔CAM_Pose"
            global PSE_T=CAM_Pose
            $ 1281 "PSE_T" "breakAfter"
            set_tcp(p[0.0,0.0,0.161,3.1415,0.0,0.0])
            movel(pose_trans(FRM_Reference, PSE_T), a=0.03, v=0.05)
          end
        end
        $ 1282 "Wait: 0.5"
        sleep(0.5)
        $ 1283 "Set"
        set_tcp(p[0.0,0.0,0.161,3.1415,0.0,0.0])
        # begin: URCap Program Node
        #   Source: SensoPart VISOR Robotic, 2.0.6, SensoPart Industriesensorik GmbH
        #   Type: VISOR Trigger
        $ 1284 "# 1 VISOR Trigger"
        visor_changeJob(1, "Object Detection Single", 6000)
        visor_trigger(1, 6000, "arm")
        # end: URCap Program Node
        $ 1285 "If visor_isResponseOk(1)"
        if ( visor_isResponseOk (1)):
          $ 1286 "CAM_CNT_Obj≔visor_partsFound(1)"
          global CAM_CNT_Obj= visor_partsFound (1)
          $ 1287 "CAM_OBJ_Pose≔visor_getPose3d(1, 0)"
          global CAM_OBJ_Pose= visor_getPose3d (1, 0)
          $ 1288 "If CAM_CNT_Obj>0"
          if (CAM_CNT_Obj>0):
            $ 1289 "CAM_OBJ_Color≔visor_getAdditionalData(1, 0)"
            global CAM_OBJ_Color= visor_getAdditionalData (1, 0)
            $ 1290 "CAM_DetectScore≔to_num(visor_getAdditionalData(1, 1))/1000"
            global CAM_DetectScore=to_num( visor_getAdditionalData (1, 1))/1000
            $ 1291 "OBJ_Detected≔ True "
            global OBJ_Detected=  True
          end
        else:
          $ 1292 "Else" "noBreak"
          $ 1293 "CAM_Captures≔CAM_Captures+1"
          global CAM_Captures=CAM_Captures+1
        end
        $ 1294 "If OBJ_Detected"
        if (OBJ_Detected):
          $ 1295 "Get object data"
          $ 1296 "PRC_CntDetect≔0"
          global PRC_CntDetect=0
          $ 1297 "Loop PRC_CntDetect<CAM_CNT_Obj"
          while (PRC_CntDetect<CAM_CNT_Obj):
            $ 1298 "get object and jig number"
            $ 1299 "If ITM_ID≟1 and JIG≟7"
            if (ITM_ID == 1  and  JIG == 7):
              $ 1300 "FRM_Reference≔FRM_Cap_SSRack"
              global FRM_Reference=FRM_Cap_SSRack
            else:
              $ 1301 "ElseIf ITM_ID≟5 and JIG≟7"
              if (ITM_ID == 5  and  JIG == 7):
                $ 1302 "FRM_Reference≔uLM_Cap_SSRack"
                global FRM_Reference=uLM_Cap_SSRack
              end
            end
            $ 1305 "PSE_T≔pose_trans(pose_inv(FRM_Reference), CAM_OBJ_Pose)"
            global PSE_T= pose_trans ( pose_inv (FRM_Reference), CAM_OBJ_Pose)
            $ 1306 "CAM_Result.append(get_pattern_counter(PSE_T, 'X', pattern=[10, 5], patternsize=[0.181, 0.081]))"
            CAM_Result.append(get_pattern_counter(PSE_T, "X", pattern=[10, 5], patternsize=[0.181, 0.081]))
            $ 1307 "PRC_CntDetect≔PRC_CntDetect+1"
            global PRC_CntDetect=PRC_CntDetect+1
          end
          $ 1308 "CAM_Done≔ True "
          global CAM_Done=  True
        else:
          $ 1309 "ElseIf CAM_Captures≥CAM_PRM_Retries"
          if (CAM_Captures >= CAM_PRM_Retries):
            $ 1310 "CAM_Done≔ True "
            global CAM_Done=  True
          else:
            $ 1311 "Else" "noBreak"
            $ 1312 "CAM_Captures≔CAM_Captures+1"
            global CAM_Captures=CAM_Captures+1
          end
        end
      end
    end
    $ 1313 "'=========='"
    # '=========='
    $ 1314 "PostSettings"
    $ 1315 "FRM_Reference≔p[0,0,0,0,0,0]"
    global FRM_Reference=p[0,0,0,0,0,0]
    $ 1316 "Set"
    set_tcp(p[0.0,0.0,0.161,3.1415,0.0,0.0])
    $ 1317 "CAM_Pose≔p[0,0,0,0,0,0]"
    global CAM_Pose=p[0,0,0,0,0,0]
    $ 1318 "Action≔0"
    global Action=0
    $ 1319 "Action_Info≔''"
    global Action_Info=""
  end
  def Sub_AMR_MiR_V3():
    $ 1320 "Sub_AMR_MiR_V3" "noBreak"
    $ 1321 "PreSettings"
    $ 1322 "AMR_TargetList≔[1,2,3,4,5,6,7,21,22,23,24,31,32,33,34,35,36,37,38,41]"
    global AMR_TargetList=[1,2,3,4,5,6,7,21,22,23,24,31,32,33,34,35,36,37,38,41]
    $ 1323 "AMR_Done≔ False "
    global AMR_Done=  False
    $ 1324 "AMR_PosActual≔T2O_Current_Pos"
    global AMR_PosActual=modbus_get_signal_status("T2O_Current_Pos")
    $ 1325 "AMR_Attemps≔T2O_Nav_Attemps"
    global AMR_Attemps=modbus_get_signal_status("T2O_Nav_Attemps")
    $ 1326 "AMR_Battery≔MiR_Battery_Lvl"
    global AMR_Battery=modbus_get_signal_status("MiR_Battery_Lvl")
    $ 1327 "AMR_Charging≔(T2O_Charging≟1)"
    global AMR_Charging=(modbus_get_signal_status("T2O_Charging") == 1)
    $ 1328 "AMR_Position≔struct(position_identifier=T2O_Current_Pos, x1=MiR_Position_X1, x2=MiR_Position_X2, y1=MiR_Position_Y1, y2=MiR_Position_Y2, theta1=MiR_Theta_1, theta2=MiR_Theta_2) "
    global AMR_Position=struct(position_identifier=modbus_get_signal_status("T2O_Current_Pos"), x1=modbus_get_signal_status("MiR_Position_X1"), x2=modbus_get_signal_status("MiR_Position_X2"), y1=modbus_get_signal_status("MiR_Position_Y1"), y2=modbus_get_signal_status("MiR_Position_Y2"), theta1=modbus_get_signal_status("MiR_Theta_1"), theta2=modbus_get_signal_status("MiR_Theta_2"))
    $ 1329 "If MiR_Mode≠7"
    if (modbus_get_signal_status("MiR_Mode") != 7):
      $ 1330 "Error"
      $ 1331 "set_error(ERROR_AMR_WRONG_MODE)"
      set_error(ERROR_AMR_WRONG_MODE)
      $ 1332 "AMR_Done≔ True "
      global AMR_Done=  True
    end
    $ 1333 "'=========='"
    # '=========='
    $ 1334 "Switch STATE"
    switch_1 = STATE
    $ 1335 "Case 1"
    if (1 == switch_1):
      $ 1336 "stopping"
      $ 1337 "If T2O_Done≟1 and O2T_Acknowledge≟0"
      if (modbus_get_signal_status("T2O_Done") == 1  and  modbus_get_signal_status("O2T_Acknowledge") == 0):
        $ 1338 "Set O2T_Acknowledge=1"
        modbus_set_output_register("O2T_Acknowledge", 1)
      end
      $ 1339 "Set MiR_CMD_Stop=On"
      modbus_set_output_signal("MiR_CMD_Stop", True)
      $ 1340 "AMR_Position.position_identifier = 0"
      AMR_Position.position_identifier = 0
      $ 1341 "AMR_Done≔ True "
      global AMR_Done=  True
    elif (2 == switch_1):
      $ 1342 "Case 2"
      $ 1343 "stopped"
      $ 1344 "If MiR_State≠3 and MiR_State≠5"
      if (modbus_get_signal_status("MiR_State") != 3  and  modbus_get_signal_status("MiR_State") != 5):
        $ 1345 "Set MiR_CMD_Stop=Off"
        modbus_set_output_signal("MiR_CMD_Stop", False)
      end
    elif (3 == switch_1):
      $ 1346 "Case 3"
      $ 1347 "resetting"
      $ 1348 "Set O2T_Mis_Main=Off"
      modbus_set_output_signal("O2T_Mis_Main", False)
      $ 1349 "Set O2T_Mis_Charge=Off"
      modbus_set_output_signal("O2T_Mis_Charge", False)
      $ 1350 "If MiR_Mis_Queue>0"
      if (modbus_get_signal_status("MiR_Mis_Queue")>0):
        $ 1351 "Set MiR_CMD_Clear_Q=On"
        modbus_set_output_signal("MiR_CMD_Clear_Q", True)
        $ 1352 "Wait MiR_Mis_Queue≟0"
        while (not(modbus_get_signal_status("MiR_Mis_Queue") == 0)):
          sync()
        end
        $ 1353 "Set MiR_CMD_Clear_Q=Off"
        modbus_set_output_signal("MiR_CMD_Clear_Q", False)
      end
      $ 1354 "If MiR_Error_ID≠0"
      if (modbus_get_signal_status("MiR_Error_ID") != 0):
        $ 1355 "Set MiR_CMD_Clear_E=On"
        modbus_set_output_signal("MiR_CMD_Clear_E", True)
        $ 1356 "Wait MiR_Error_ID≟0"
        while (not(modbus_get_signal_status("MiR_Error_ID") == 0)):
          sync()
        end
        $ 1357 "Set MiR_CMD_Clear_E=Off"
        modbus_set_output_signal("MiR_CMD_Clear_E", False)
      end
      $ 1358 "Set O2T_Action=0"
      modbus_set_output_register("O2T_Action", 0)
      $ 1359 "Set O2T_Acknowledge=0"
      modbus_set_output_register("O2T_Acknowledge", 0)
      $ 1360 "Set O2T_Target_Pos=0"
      modbus_set_output_register("O2T_Target_Pos", 0)
      $ 1361 "Set O2T_Footprint=0"
      modbus_set_output_register("O2T_Footprint", 0)
      $ 1362 "Set O2T_ProtectOff=0"
      modbus_set_output_register("O2T_ProtectOff", 0)
      $ 1363 "Set O2T_Dock=0"
      modbus_set_output_register("O2T_Dock", 0)
      $ 1364 "AMR_Attemps≔0"
      global AMR_Attemps=0
      $ 1365 "AMR_PosTarget≔0"
      global AMR_PosTarget=0
      $ 1366 "AMR_Step≔0"
      global AMR_Step=0
      $ 1367 "AMR_AtTarget≔ False "
      global AMR_AtTarget=  False
      $ 1368 "If MiR_State≟4 or MiR_State≟3 or MiR_State≟10"
      if (modbus_get_signal_status("MiR_State") == 4  or  modbus_get_signal_status("MiR_State") == 3  or  modbus_get_signal_status("MiR_State") == 10):
        $ 1369 "AMR_Done≔ True "
        global AMR_Done=  True
      end
    elif (5 == switch_1):
      $ 1370 "Case 5"
      $ 1371 "starting"
      $ 1372 "If MiR_State≟4"
      if (modbus_get_signal_status("MiR_State") == 4):
        $ 1373 "Set MiR_CMD_Start=On"
        modbus_set_output_signal("MiR_CMD_Start", True)
        $ 1374 "Wait MiR_State≠4"
        while (not(modbus_get_signal_status("MiR_State") != 4)):
          sync()
        end
        $ 1375 "Set MiR_CMD_Start=Off"
        modbus_set_output_signal("MiR_CMD_Start", False)
        $ 1376 "AMR_Done≔ True "
        global AMR_Done=  True
      else:
        $ 1377 "ElseIf MiR_State≟10"
        if (modbus_get_signal_status("MiR_State") == 10):
          $ 1378 "'MiR in protective stop. Wait'"
          # 'MiR in protective stop. Wait'
          $ 1379 "AMR_Done≔ True "
          global AMR_Done=  True
        else:
          $ 1380 "ElseIf MiR_State≟3"
          if (modbus_get_signal_status("MiR_State") == 3):
            $ 1381 "AMR_Done≔ True "
            global AMR_Done=  True
          end
        end
      end
    elif (6 == switch_1):
      $ 1382 "Case 6"
      $ 1383 "execute"
      $ 1384 "AMR_AtTarget≔(AMR_PosActual≟AMR_PosTarget)"
      global AMR_AtTarget=(AMR_PosActual == AMR_PosTarget)
      $ 1385 "Switch AMR_Step"
      switch_2 = AMR_Step
      $ 1386 "Case 0"
      if (0 == switch_2):
        $ 1387 "If  not AMR_AtTarget"
        if (  not  AMR_AtTarget):
          $ 1388 "AMR_Step≔1"
          global AMR_Step=1
        else:
          $ 1389 "Else" "noBreak"
          $ 1390 "AMR_Done≔ True "
          global AMR_Done=  True
        end
      elif (1 == switch_2):
        $ 1391 "Case 1"
        $ 1392 "general Settings"
        $ 1393 "Set O2T_Acknowledge=0"
        modbus_set_output_register("O2T_Acknowledge", 0)
        $ 1394 "check for error"
        $ 1395 "If OBJ_Picked and MiR_State≟10"
        if (OBJ_Picked  and  modbus_get_signal_status("MiR_State") == 10):
          $ 1396 "Error"
          $ 1397 "set_error(ERROR_ROBOT_ARM_NOT_IN_HOME_POSE)"
          set_error(ERROR_ROBOT_ARM_NOT_IN_HOME_POSE)
          $ 1398 "Action≔0"
          global Action=0
        else:
          $ 1399 "ElseIf  not found_in_list(AMR_PosTarget, AMR_TargetList)"
          if (  not  found_in_list(AMR_PosTarget, AMR_TargetList)):
            $ 1400 "Error"
            $ 1401 "set_error(ERROR_UNKNOWN_POSE)"
            set_error(ERROR_UNKNOWN_POSE)
            $ 1402 "Action≔0"
            global Action=0
          end
        end
        $ 1403 "If MiR_State≟3"
        if (modbus_get_signal_status("MiR_State") == 3):
          $ 1404 "Set MiR_CMD_Start=Off"
          modbus_set_output_signal("MiR_CMD_Start", False)
          $ 1405 "Switch Action"
          switch_3 = Action
          $ 1406 "Case 51"
          if (51 == switch_3):
            $ 1407 "Charge"
            $ 1408 "'trigger the charging mission'"
            # 'trigger the charging mission'
            $ 1409 "'target pos is predefined'"
            # 'target pos is predefined'
            $ 1410 "Set O2T_Footprint=0"
            modbus_set_output_register("O2T_Footprint", 0)
            $ 1411 "Set O2T_Action=1"
            modbus_set_output_register("O2T_Action", 1)
            $ 1412 "If MiR_Mis_Queue≟0"
            if (modbus_get_signal_status("MiR_Mis_Queue") == 0):
              $ 1413 "Set O2T_Mis_Charge=On"
              modbus_set_output_signal("O2T_Mis_Charge", True)
              $ 1414 "Wait MiR_Mis_Queue≥1"
              while (not(modbus_get_signal_status("MiR_Mis_Queue") >= 1)):
                sync()
              end
              $ 1415 "Set O2T_Mis_Charge=Off"
              modbus_set_output_signal("O2T_Mis_Charge", False)
            end
          elif (52 == switch_3):
            $ 1416 "Case 52"
            $ 1417 "Navigate"
            $ 1418 "'trigger the standard missoin'"
            # 'trigger the standard missoin'
            $ 1419 "Set O2T_Footprint=AMR_FootprintID"
            modbus_set_output_register("O2T_Footprint", AMR_FootprintID)
            $ 1420 "Set O2T_Target_Pos=AMR_PosTarget"
            modbus_set_output_register("O2T_Target_Pos", AMR_PosTarget)
            $ 1421 "Set O2T_Action=2"
            modbus_set_output_register("O2T_Action", 2)
            $ 1422 "If MiR_Mis_Queue≟0"
            if (modbus_get_signal_status("MiR_Mis_Queue") == 0):
              $ 1423 "Set O2T_Mis_Main=On"
              modbus_set_output_signal("O2T_Mis_Main", True)
              $ 1424 "Wait MiR_Mis_Queue≥1"
              while (not(modbus_get_signal_status("MiR_Mis_Queue") >= 1)):
                sync()
              end
              $ 1425 "Set O2T_Mis_Main=Off"
              modbus_set_output_signal("O2T_Mis_Main", False)
            end
          end
        else:
          $ 1426 "ElseIf MiR_State≟4"
          if (modbus_get_signal_status("MiR_State") == 4):
            $ 1427 "Set MiR_CMD_Start=On"
            modbus_set_output_signal("MiR_CMD_Start", True)
          else:
            $ 1428 "ElseIf MiR_State≟5"
            if (modbus_get_signal_status("MiR_State") == 5):
              $ 1429 "AMR_Step≔2"
              global AMR_Step=2
            else:
              $ 1430 "ElseIf MiR_State≟10"
              if (modbus_get_signal_status("MiR_State") == 10):
                $ 1431 "'AMR still in safeguard stop'"
                # 'AMR still in safeguard stop'
              end
            end
          end
        end
      elif (2 == switch_2):
        $ 1432 "Case 2"
        $ 1433 "acknowledge handshake"
        $ 1434 "If T2O_Done≟1 and O2T_Acknowledge≟0"
        if (modbus_get_signal_status("T2O_Done") == 1  and  modbus_get_signal_status("O2T_Acknowledge") == 0):
          $ 1435 "Set O2T_Acknowledge=1"
          modbus_set_output_register("O2T_Acknowledge", 1)
        else:
          $ 1436 "ElseIf T2O_Done≟0 and O2T_Acknowledge≟1"
          if (modbus_get_signal_status("T2O_Done") == 0  and  modbus_get_signal_status("O2T_Acknowledge") == 1):
            $ 1437 "Set O2T_Acknowledge=0"
            modbus_set_output_register("O2T_Acknowledge", 0)
            $ 1438 "AMR_AtTarget≔(AMR_PosActual≟AMR_PosTarget)"
            global AMR_AtTarget=(AMR_PosActual == AMR_PosTarget)
            $ 1439 "AMR_Done≔ True "
            global AMR_Done=  True
          end
        end
      end
      $ 1440 "translate errors"
      $ 1441 "If AMR_Done"
      if (AMR_Done):
        $ 1442 "Switch T2O_Error_ID"
        switch_2 = modbus_get_signal_status("T2O_Error_ID")
        $ 1443 "Case 2003"
        if (2003 == switch_2):
          $ 1444 "error"
          $ 1445 "set_error(ERROR_NOT_DOCKED)"
          set_error(ERROR_NOT_DOCKED)
        elif (2007 == switch_2):
          $ 1446 "Case 2007"
          $ 1447 "error"
          $ 1448 "set_error(ERROR_NOT_REACHABLE_TARGET)"
          set_error(ERROR_NOT_REACHABLE_TARGET)
        elif (2008 == switch_2):
          $ 1449 "Case 2008"
          $ 1450 "error"
          $ 1451 "set_error(ERROR_CHARGING_NOT_STARTED)"
          set_error(ERROR_CHARGING_NOT_STARTED)
        end
      end
    elif (7 == switch_1):
      $ 1452 "Case 7"
      $ 1453 "completing"
      $ 1454 "If MiR_Mis_Queue>0"
      if (modbus_get_signal_status("MiR_Mis_Queue")>0):
        $ 1455 "Set MiR_CMD_Abort=On"
        modbus_set_output_signal("MiR_CMD_Abort", True)
        $ 1456 "Wait MiR_Mis_Queue≟0"
        while (not(modbus_get_signal_status("MiR_Mis_Queue") == 0)):
          sync()
        end
        $ 1457 "Set MiR_CMD_Abort=Off"
        modbus_set_output_signal("MiR_CMD_Abort", False)
      end
      $ 1458 "If MiR_State≟3 or MiR_State≟10"
      if (modbus_get_signal_status("MiR_State") == 3  or  modbus_get_signal_status("MiR_State") == 10):
        $ 1459 "AMR_Done≔ True "
        global AMR_Done=  True
      end
    elif (9 == switch_1):
      $ 1460 "Case 9"
      $ 1461 "holding"
      $ 1462 "Set MiR_CMD_Abort=On"
      modbus_set_output_signal("MiR_CMD_Abort", True)
      $ 1463 "If MiR_State≟3 or MiR_State≟10"
      if (modbus_get_signal_status("MiR_State") == 3  or  modbus_get_signal_status("MiR_State") == 10):
        $ 1464 "Set MiR_CMD_Abort=Off"
        modbus_set_output_signal("MiR_CMD_Abort", False)
        $ 1465 "AMR_Done≔ True "
        global AMR_Done=  True
      end
    elif (11 == switch_1):
      $ 1466 "Case 11"
      $ 1467 "unholding"
      $ 1468 "Set MiR_CMD_Start=On"
      modbus_set_output_signal("MiR_CMD_Start", True)
      $ 1469 "If MiR_State≠4"
      if (modbus_get_signal_status("MiR_State") != 4):
        $ 1470 "Set MiR_CMD_Start=Off"
        modbus_set_output_signal("MiR_CMD_Start", False)
        $ 1471 "AMR_Step≔0"
        global AMR_Step=0
        $ 1472 "AMR_Done≔ True "
        global AMR_Done=  True
      end
    elif (12 == switch_1):
      $ 1473 "Case 12"
      $ 1474 "suspending"
      $ 1475 "'none'"
      # 'none'
    elif (14 == switch_1):
      $ 1476 "Case 14"
      $ 1477 "unsuspending"
      $ 1478 "'none'"
      # 'none'
    elif (15 == switch_1):
      $ 1479 "Case 15"
      $ 1480 "aborting"
      $ 1481 "Set MiR_CMD_Abort=On"
      modbus_set_output_signal("MiR_CMD_Abort", True)
      $ 1482 "Wait MiR_State≟3"
      while (not(modbus_get_signal_status("MiR_State") == 3)):
        sync()
      end
      $ 1483 "Set MiR_CMD_Abort=Off"
      modbus_set_output_signal("MiR_CMD_Abort", False)
    elif (17 == switch_1):
      $ 1484 "Case 17"
      $ 1485 "clearing"
      $ 1486 "If MiR_Error_ID≠0"
      if (modbus_get_signal_status("MiR_Error_ID") != 0):
        $ 1487 "Set MiR_CMD_Clear_E=On"
        modbus_set_output_signal("MiR_CMD_Clear_E", True)
        $ 1488 "Wait MiR_Error_ID≟0"
        while (not(modbus_get_signal_status("MiR_Error_ID") == 0)):
          sync()
        end
        $ 1489 "Set MiR_CMD_Clear_E=Off"
        modbus_set_output_signal("MiR_CMD_Clear_E", False)
      end
      $ 1490 "If MiR_Error_ID≟0"
      if (modbus_get_signal_status("MiR_Error_ID") == 0):
        $ 1491 "AMR_Done≔ True "
        global AMR_Done=  True
      end
    end
    $ 1492 "'=========='"
    # '=========='
    $ 1493 "PostSettings"
    $ 1494 "AMR_Position≔struct(position_identifier=T2O_Current_Pos, x1=MiR_Position_X1, x2=MiR_Position_X2, y1=MiR_Position_Y1, y2=MiR_Position_Y2, theta1=MiR_Theta_1, theta2=MiR_Theta_2) "
    global AMR_Position=struct(position_identifier=modbus_get_signal_status("T2O_Current_Pos"), x1=modbus_get_signal_status("MiR_Position_X1"), x2=modbus_get_signal_status("MiR_Position_X2"), y1=modbus_get_signal_status("MiR_Position_Y1"), y2=modbus_get_signal_status("MiR_Position_Y2"), theta1=modbus_get_signal_status("MiR_Theta_1"), theta2=modbus_get_signal_status("MiR_Theta_2"))
  end
  def Sub_Action_V4():
    $ 1495 "Sub_Action_V4" "noBreak"
    $ 1496 "PreSettings"
    $ 1497 "init poses"
    $ 1498 "PSE_A≔p[0,0,0,0,0,0]"
    global PSE_A=p[0,0,0,0,0,0]
    $ 1499 "PSE_A_H≔p[0,0,0,0,0,0]"
    global PSE_A_H=p[0,0,0,0,0,0]
    $ 1500 "PSE_T≔p[0,0,0,0,0,0]"
    global PSE_T=p[0,0,0,0,0,0]
    $ 1501 "PSE_T_H≔p[0,0,0,0,0,0]"
    global PSE_T_H=p[0,0,0,0,0,0]
    $ 1502 "PSE_G≔p[0,0,0,0,0,0]"
    global PSE_G=p[0,0,0,0,0,0]
    $ 1503 "PSE_G_H≔p[0,0,0,0,0,0]"
    global PSE_G_H=p[0,0,0,0,0,0]
    $ 1504 "PSE_R≔p[0,0,0,0,0,0]"
    global PSE_R=p[0,0,0,0,0,0]
    $ 1505 "PSE_R_H≔p[0,0,0,0,0,0]"
    global PSE_R_H=p[0,0,0,0,0,0]
    $ 1506 "JNT_Q≔[0,0,0,0,0,0]"
    global JNT_Q=[0,0,0,0,0,0]
    $ 1507 "JNT_S≔[0,0,0,0,0,0]"
    global JNT_S=[0,0,0,0,0,0]
    $ 1508 "Gripping parameters"
    $ 1509 "OBJ = find_object_by_type(OBJs, OBJ_Type)"
    OBJ = find_object_by_type(OBJs, OBJ_Type)
    $ 1510 "GRP_Open_Pos≔OBJ.dimension.diameter * 1000 + 6"
    global GRP_Open_Pos=OBJ.dimension.diameter * 1000 + 6
    $ 1511 "GRP_Offset≔OBJ.gripper_offset"
    global GRP_Offset=OBJ.gripper_offset
    $ 1512 "rq_set_force_norm(50)"
     rq_set_force_norm (50)
    $ 1513 "rq_set_speed_norm(50)"
     rq_set_speed_norm (50)
    $ 1514 "Switch ITM_ID"
    switch_1 = ITM_ID
    $ 1515 "Case 1"
    if (1 == switch_1):
      $ 1516 "uML"
      $ 1517 "JIG2 = find_object_by_type(JIGs, JIG)"
      JIG2 = find_object_by_type(JIGs, JIG)
      $ 1518 "JIG_Offset≔JIG2.jig_offset"
      global JIG_Offset=JIG2.jig_offset
      $ 1519 "Switch JIG"
      switch_2 = JIG
      $ 1520 "Case 1"
      if (1 == switch_2):
        $ 1521 "3FG"
        $ 1522 "define poses"
        $ 1523 "FRM_Reference≔ULM_3FG"
        global FRM_Reference=ULM_3FG
        $ 1524 "JNT_Q≔JNT_HOME"
        global JNT_Q=JNT_HOME
        $ 1525 "PSE_T≔pose_trans(GRP_Offset, JIG_Offset)"
        global PSE_T= pose_trans (GRP_Offset, JIG_Offset)
        $ 1526 "PSE_A≔pose_trans(PSE_T, p[0,0,0.100,0,0,0])"
        global PSE_A= pose_trans (PSE_T, p[0,0,0.100,0,0,0])
        $ 1527 "PSE_R≔pose_add(PSE_T, p[0,0,0.100,0,0,0])"
        global PSE_R= pose_add (PSE_T, p[0,0,0.100,0,0,0])
      elif (2 == switch_2):
        $ 1528 "Case 2"
        $ 1529 "Input"
        $ 1530 "'CHANGE THE REFERENCE TO THE FRAME TO MOVE IN'"
        # 'CHANGE THE REFERENCE TO THE FRAME TO MOVE IN'
        $ 1531 "define poses"
        $ 1532 "FRM_Reference≔ULM_Input"
        global FRM_Reference=ULM_Input
        $ 1533 "PSE_T≔pose_trans(pose_trans(get_pattern_pos_rectangle(OBJ_Nbr, 'X', [10,5], patternsize=[0.181,0.081]), GRP_Offset), JIG_Offset)"
        global PSE_T= pose_trans ( pose_trans (get_pattern_pos_rectangle(OBJ_Nbr, "X", [10,5], patternsize=[0.181,0.081]), GRP_Offset), JIG_Offset)
        $ 1534 "If Action≟1"
        if (Action == 1):
          $ 1535 "PSE_R≔pose_add(PSE_T, p[0,0,0.200,0,0,0])"
          global PSE_R= pose_add (PSE_T, p[0,0,0.200,0,0,0])
          $ 1536 "PSE_A≔pose_add(PSE_T, p[0,0,0.100,0,0,0])"
          global PSE_A= pose_add (PSE_T, p[0,0,0.100,0,0,0])
        else:
          $ 1537 "ElseIf Action≟2"
          if (Action == 2):
            $ 1538 "PSE_R≔pose_add(PSE_T, p[0,0,0.100,0,0,0])"
            global PSE_R= pose_add (PSE_T, p[0,0,0.100,0,0,0])
            $ 1539 "PSE_A≔pose_add(PSE_T, p[0,0,0.200,0,0,0])"
            global PSE_A= pose_add (PSE_T, p[0,0,0.200,0,0,0])
          end
        end
      elif (3 == switch_2):
        $ 1540 "Case 3"
        $ 1541 "Output"
        $ 1542 "'CHANGE THE REFERENCE TO THE FRAME TO MOVE IN'"
        # 'CHANGE THE REFERENCE TO THE FRAME TO MOVE IN'
        $ 1543 "define poses"
        $ 1544 "FRM_Reference≔ULM_Output"
        global FRM_Reference=ULM_Output
        $ 1545 "PSE_T≔pose_trans(pose_trans(get_pattern_pos_rectangle(OBJ_Nbr, 'X', [10,5], patternsize=[0.181,0.081]), GRP_Offset), JIG_Offset)"
        global PSE_T= pose_trans ( pose_trans (get_pattern_pos_rectangle(OBJ_Nbr, "X", [10,5], patternsize=[0.181,0.081]), GRP_Offset), JIG_Offset)
        $ 1547 "If Action≟1"
        if (Action == 1):
          $ 1548 "PSE_R≔pose_add(PSE_T, p[0,0,0.200,0,0,0])"
          global PSE_R= pose_add (PSE_T, p[0,0,0.200,0,0,0])
          $ 1549 "PSE_A≔pose_add(PSE_T, p[0,0,0.100,0,0,0])"
          global PSE_A= pose_add (PSE_T, p[0,0,0.100,0,0,0])
        else:
          $ 1550 "ElseIf Action≟2"
          if (Action == 2):
            $ 1551 "PSE_R≔pose_add(PSE_T, p[0,0,0.100,0,0,0])"
            global PSE_R= pose_add (PSE_T, p[0,0,0.100,0,0,0])
            $ 1552 "PSE_A≔pose_add(PSE_T, p[0,0,0.200,0,0,0])"
            global PSE_A= pose_add (PSE_T, p[0,0,0.200,0,0,0])
          end
        end
      elif (4 == switch_2):
        $ 1553 "Case 4"
        $ 1554 "jig centrifuge racks"
        $ 1555 "define poses"
        $ 1556 "FRM_Reference≔ULM_Cent_Racks"
        global FRM_Reference=ULM_Cent_Racks
        $ 1557 "PSE_T≔get_pattern_pos_rectangle(JIG_Slot, 'X', [4,1], patternsize=[0.291,0])"
        global PSE_T=get_pattern_pos_rectangle(JIG_Slot, "X", [4,1], patternsize=[0.291,0])
        $ 1558 "If OBJ_Nbr≠0"
        if (OBJ_Nbr != 0):
          $ 1559 "PSE_T≔pose_trans(pose_trans(PSE_T, get_pattern_pos_rectangle(OBJ_Nbr, 'X', [3,3], patternsize=[0.060,0.060])),p[-0.030, -0.030,0,0,0,3.927])"
          global PSE_T= pose_trans ( pose_trans (PSE_T, get_pattern_pos_rectangle(OBJ_Nbr, "X", [3,3], patternsize=[0.060,0.060])),p[-0.030, -0.030,0,0,0,3.927])
        end
        $ 1560 "PSE_T≔pose_trans(PSE_T, GRP_Offset)"
        global PSE_T= pose_trans (PSE_T, GRP_Offset)
        $ 1561 "If Action≟1"
        if (Action == 1):
          $ 1562 "PSE_R≔pose_add(PSE_T, p[0,0,0.200,0,0,0])"
          global PSE_R= pose_add (PSE_T, p[0,0,0.200,0,0,0])
          $ 1563 "PSE_A≔pose_add(PSE_T, p[0,0,0.100,0,0,0])"
          global PSE_A= pose_add (PSE_T, p[0,0,0.100,0,0,0])
        else:
          $ 1564 "ElseIf Action≟2"
          if (Action == 2):
            $ 1565 "PSE_R≔pose_add(PSE_T, p[0,0,0.100,0,0,0])"
            global PSE_R= pose_add (PSE_T, p[0,0,0.100,0,0,0])
            $ 1566 "PSE_A≔pose_add(PSE_T, p[0,0,0.200,0,0,0])"
            global PSE_A= pose_add (PSE_T, p[0,0,0.200,0,0,0])
          end
        end
      elif (6 == switch_2):
        $ 1567 "Case 6"
        $ 1568 "Caps bin"
        $ 1569 "define poses"
        $ 1570 "'Drop cap'"
        # 'Drop cap'
        $ 1571 "FRM_Reference=ULM_Cap_Bin"
        FRM_Reference=ULM_Cap_Bin
        $ 1572 "PSE_T≔pose_RPY2RotVec(p[0,0,0,0,0,0])"
        global PSE_T=pose_RPY2RotVec(p[0,0,0,0,0,0])
        $ 1573 "PSE_T_H≔pose_add(PSE_T, p[0,0,-0.011,0,0,0])"
        global PSE_T_H= pose_add (PSE_T, p[0,0,-0.011,0,0,0])
        $ 1574 "PSE_A≔pose_trans(PSE_T, p[0,0,0.1,0,0,0])"
        global PSE_A= pose_trans (PSE_T, p[0,0,0.1,0,0,0])
        $ 1575 "PSE_R_H≔pose_add(PSE_T, p[0,0,0.100,0,0,0])"
        global PSE_R_H= pose_add (PSE_T, p[0,0,0.100,0,0,0])
        $ 1576 "PSE_R≔pose_add(PSE_T, p[0,0,0.100,0,0,0])"
        global PSE_R= pose_add (PSE_T, p[0,0,0.100,0,0,0])
      elif (7 == switch_2):
        $ 1577 "Case 7"
      elif (8 == switch_2):
        $ 1602 "Case 8"
        $ 1603 "NoK"
        $ 1604 "define poses"
        $ 1605 "'NoK'"
        # 'NoK'
        $ 1606 "FRM_Reference=ULM_NoK"
        FRM_Reference=ULM_NoK
        $ 1607 "PSE_T≔pose_RPY2RotVec(p[0,0,0,0,0,0])"
        global PSE_T=pose_RPY2RotVec(p[0,0,0,0,0,0])
        $ 1608 "PSE_A≔pose_trans(PSE_T, p[0,0,0.1,0,0,0])"
        global PSE_A= pose_trans (PSE_T, p[0,0,0.1,0,0,0])
        $ 1609 "PSE_R≔pose_add(PSE_T, p[0,0,0.100,0,0,0])"
        global PSE_R= pose_add (PSE_T, p[0,0,0.100,0,0,0])
      elif (9 == switch_2):
        $ 1610 "Case 9"
      elif (10 == switch_2):
        $ 1618 "Case 10"
      elif (11 == switch_2):
        $ 1626 "Case 11"
      elif (12 == switch_2):
        $ 1634 "Case 12"
      end
    elif (2 == switch_1):
      $ 1642 "Case 2"
      $ 1643 "Centrifuge"
      $ 1644 "'CHANGE THE REFERENCE TO THE FRAME TO MOVE IN'"
      # 'CHANGE THE REFERENCE TO THE FRAME TO MOVE IN'
      $ 1645 "define poses"
      $ 1646 "FRM_Reference≔FRM_Centrifuge"
      global FRM_Reference=FRM_Centrifuge
      $ 1647 "PSE_T≔GRP_Offset"
      global PSE_T=GRP_Offset
      $ 1648 "If Action≟8"
      if (Action == 8):
        $ 1649 "PSE_R≔pose_add(PSE_T, p[0,0,0.250,0,0,0])"
        global PSE_R= pose_add (PSE_T, p[0,0,0.250,0,0,0])
        $ 1650 "PSE_A≔pose_add(PSE_T, p[0,0,0.150,0,0,0])"
        global PSE_A= pose_add (PSE_T, p[0,0,0.150,0,0,0])
      else:
        $ 1651 "ElseIf Action≟7"
        if (Action == 7):
          $ 1652 "PSE_R≔pose_add(PSE_T, p[0,0,0.150,0,0,0])"
          global PSE_R= pose_add (PSE_T, p[0,0,0.150,0,0,0])
          $ 1653 "PSE_A≔pose_add(PSE_T, p[0,0,0.250,0,0,0])"
          global PSE_A= pose_add (PSE_T, p[0,0,0.250,0,0,0])
        end
      end
    elif (3 == switch_1):
      $ 1654 "Case 3"
      $ 1655 "Output"
      $ 1656 "'CHANGE THE REFERENCE TO THE FRAME TO MOVE IN'"
      # 'CHANGE THE REFERENCE TO THE FRAME TO MOVE IN'
      $ 1657 "define poses"
      $ 1658 "FRM_Reference≔Base_const"
      global FRM_Reference=p[0.0,0.0,0.0,0.0,0.0,0.0]
      $ 1659 "PSE_T≔p[0,0,0,0,0,0]"
      global PSE_T=p[0,0,0,0,0,0]
      $ 1660 "PSE_A≔pose_add(PSE_T, p[0,0,0.150,0,0,0])"
      global PSE_A= pose_add (PSE_T, p[0,0,0.150,0,0,0])
      $ 1661 "PSE_R≔pose_add(PSE_T, p[0,0,0.100,0,0,0])"
      global PSE_R= pose_add (PSE_T, p[0,0,0.100,0,0,0])
    elif (5 == switch_1):
      $ 1662 "Case 5"
      $ 1663 "Sarstedt Pickup Table"
      $ 1664 "'CHANGE THE REFERENCE TO THE FRAME TO MOVE IN'"
      # 'CHANGE THE REFERENCE TO THE FRAME TO MOVE IN'
      $ 1665 "Switch JIG"
      switch_2 = JIG
      $ 1666 "Case 7"
      if (7 == switch_2):
        $ 1679 "Sarstedt"
        $ 1680 "'CHANGE THE REFERENCE TO THE FRAME TO MOVE IN'"
        # 'CHANGE THE REFERENCE TO THE FRAME TO MOVE IN'
        $ 1686 "If TASK.ID≟10"
        if (TASK.ID == 10):
          $ 1687 "Frame & Position Params"
          $ 1688 "FRM_Reference = CAM_LM_SSRack"
          FRM_Reference = CAM_LM_SSRack
          $ 1689 "PSE_T≔uLM_SS_PickPlc"
          global PSE_T=uLM_SS_PickPlc
          $ 1690 "PSE_A≔pose_trans(PSE_T, p[0,0,0.1,0,0,0])"
          global PSE_A= pose_trans (PSE_T, p[0,0,0.1,0,0,0])
          $ 1691 "PSE_R≔pose_add(PSE_T, p[0,0,0.1,0,0,0])"
          global PSE_R= pose_add (PSE_T, p[0,0,0.1,0,0,0])
        end
      end
    elif (13 == switch_1):
      $ 1698 "Case 13"
      $ 1699 "Sarstedt Pickup Table"
      $ 1700 "'CHANGE THE REFERENCE TO THE FRAME TO MOVE IN'"
      # 'CHANGE THE REFERENCE TO THE FRAME TO MOVE IN'
      $ 1701 "Switch JIG"
      switch_2 = JIG
      $ 1702 "Case 7"
      if (7 == switch_2):
        $ 1715 "Bottle"
        $ 1716 "'CHANGE THE REFERENCE TO THE FRAME TO MOVE IN'"
        # 'CHANGE THE REFERENCE TO THE FRAME TO MOVE IN'
        $ 1722 "If TASK.ID≟43"
        if (TASK.ID == 43):
          $ 1723 "Frame & Position Params"
          $ 1725 "PSE_T≔uLM_SS_PickPlc"
          global PSE_T=uLM_SS_PickPlc
          $ 1726 "PSE_A≔pose_trans(PSE_T, p[0,0,0.1,0,0,0])"
          global PSE_A= pose_trans (PSE_T, p[0,0,0.1,0,0,0])
          $ 1727 "PSE_R≔pose_add(PSE_T, p[0,0,0.1,0,0,0])"
          global PSE_R= pose_add (PSE_T, p[0,0,0.1,0,0,0])
        end
      end
    end
    $ 1734 "Additional check"
    $ 1735 "If  not is_reachable(FRM_Reference,[PSE_A,PSE_A_H,PSE_T,PSE_T_H,PSE_R,PSE_R_H])"
    if (  not  is_reachable(FRM_Reference,[PSE_A,PSE_A_H,PSE_T,PSE_T_H,PSE_R,PSE_R_H])):
      $ 1736 "Error"
      $ 1737 "set_error(ERROR_POSE_NOT_REACHABLE)"
      set_error(ERROR_POSE_NOT_REACHABLE)
      $ 1738 "Action≔0"
      global Action=0
    end
    $ 1739 "'=========='"
    # '=========='
    $ 1740 "Switch Action"
    switch_1 = Action
    $ 1741 "Case 1"
    if (1 == switch_1):
      $ 1742 "Pick"
      $ 1743 "Action_Info≔'pick object'"
      global Action_Info="pick object"
      $ 1744 "do_transition(pose_trans(FRM_Reference, PSE_T), keep_rxry=OBJ_Picked)"
      do_transition( pose_trans (FRM_Reference, PSE_T), keep_rxry=OBJ_Picked)
      $ 1745 "EOAT"
      $ 1746 "If  not OBJ_Picked"
      if (  not  OBJ_Picked):
        $ 1747 "rq_move_and_wait_mm(GRP_Open_Pos)"
         rq_move_and_wait_mm (GRP_Open_Pos)
      end
      $ 1748 "If PSE_A_H≠PSE_Z"
      if (PSE_A_H != PSE_Z):
        $ 1749 "If JNT_Q≠JNT_Z"
        if (JNT_Q != JNT_Z):
          $ 1750 "movej(get_inverse_kin(pose_trans(FRM_Reference, PSE_A_H), qnear=JNT_Q), r=0.050)"
          movej(get_inverse_kin( pose_trans (FRM_Reference, PSE_A_H), qnear=JNT_Q), r=0.050)
        else:
          $ 1751 "Else" "noBreak"
          $ 1752 "movej(pose_trans(FRM_Reference, PSE_A_H), r=0.050)"
          movej( pose_trans (FRM_Reference, PSE_A_H), r=0.050)
        end
      end
      $ 1753 "If PSE_A≠PSE_Z"
      if (PSE_A != PSE_Z):
        $ 1754 "If JNT_Q≠JNT_Z"
        if (JNT_Q != JNT_Z):
          $ 1755 "movej(get_inverse_kin(pose_trans(FRM_Reference, PSE_A), qnear=JNT_Q), r=0.020)"
          movej(get_inverse_kin( pose_trans (FRM_Reference, PSE_A), qnear=JNT_Q), r=0.020)
        else:
          $ 1756 "Else" "noBreak"
          $ 1757 "movej(pose_trans(FRM_Reference, PSE_A), r=0.020)"
          movej( pose_trans (FRM_Reference, PSE_A), r=0.020)
        end
      end
      $ 1758 "MoveL"
      $ 1759 "If PSE_T_H≠PSE_Z"
      if (PSE_T_H != PSE_Z):
        $ 1760 "PSE_T_H" "breakAfter"
        movel(pose_trans(FRM_Reference, PSE_T_H), a=0.5, v=0.4, r=0.01)
      end
      $ 1761 "PSE_T" "breakAfter"
      movel(pose_trans(FRM_Reference, PSE_T), a=0.08, v=0.12)
      $ 1762 "EOAT"
      $ 1763 "rq_set_force_norm(50)"
       rq_set_force_norm (50)
      $ 1764 "rq_close_and_wait()"
       rq_close_and_wait ()
      $ 1765 "OBJ_Picked≔rq_is_object_detected()"
      global OBJ_Picked= rq_is_object_detected ()
      $ 1766 "If  not OBJ_Picked"
      if (  not  OBJ_Picked):
        $ 1767 "set_error(ERROR_NO_OBJECT_TO_PICK)"
        set_error(ERROR_NO_OBJECT_TO_PICK)
      end
      $ 1768 "EXTT"
      $ 1769 "Switch JIG"
      switch_2 = JIG
      $ 1770 "Case 1"
      if (1 == switch_2):
        $ 1771 "3FG"
        $ 1772 "If OBJ_Picked"
        if (OBJ_Picked):
          $ 1773 "Set GRP_3F_Open=On"
          set_standard_digital_out(5, True)
        end
      end
      $ 1774 "If PSE_R_H≠PSE_Z"
      if (PSE_R_H != PSE_Z):
        $ 1775 "PSE_R" "breakAfter"
        movel(pose_trans(FRM_Reference, PSE_R), a=0.5, v=0.4, r=0.01)
        $ 1776 "PSE_R_H" "breakAfter"
        movel(pose_trans(FRM_Reference, PSE_R_H), a=0.5, v=0.4)
      else:
        $ 1777 "Else" "noBreak"
        $ 1778 "PSE_R" "breakAfter"
        movel(pose_trans(FRM_Reference, PSE_R), a=0.5, v=0.4)
      end
    elif (2 == switch_1):
      $ 1779 "Case 2"
      $ 1780 "Place"
      $ 1781 "Action_Info≔'place object'"
      global Action_Info="place object"
      $ 1782 "do_transition(pose_trans(FRM_Reference, PSE_T), keep_rxry=OBJ_Picked)"
      do_transition( pose_trans (FRM_Reference, PSE_T), keep_rxry=OBJ_Picked)
      $ 1783 "EXTT"
      $ 1784 "Switch JIG"
      switch_2 = JIG
      $ 1785 "Case 1"
      if (1 == switch_2):
        $ 1786 "3FG"
        $ 1787 "If OBJ_Picked"
        if (OBJ_Picked):
          $ 1788 "Set GRP_3F_Open=On"
          set_standard_digital_out(5, True)
        end
      end
      $ 1789 "If PSE_A_H≠PSE_Z"
      if (PSE_A_H != PSE_Z):
        $ 1790 "If JNT_Q≠JNT_Z"
        if (JNT_Q != JNT_Z):
          $ 1791 "movej(get_inverse_kin(pose_trans(FRM_Reference, PSE_A_H), qnear=JNT_Q), r=0.050)"
          movej(get_inverse_kin( pose_trans (FRM_Reference, PSE_A_H), qnear=JNT_Q), r=0.050)
        else:
          $ 1792 "Else" "noBreak"
          $ 1793 "movej(pose_trans(FRM_Reference, PSE_A_H), r=0.050)"
          movej( pose_trans (FRM_Reference, PSE_A_H), r=0.050)
        end
      end
      $ 1794 "If PSE_A≠PSE_Z"
      if (PSE_A != PSE_Z):
        $ 1795 "If JNT_Q≠JNT_Z"
        if (JNT_Q != JNT_Z):
          $ 1796 "movej(get_inverse_kin(pose_trans(FRM_Reference, PSE_A), qnear=JNT_Q), r=0.020)"
          movej(get_inverse_kin( pose_trans (FRM_Reference, PSE_A), qnear=JNT_Q), r=0.020)
        else:
          $ 1797 "Else" "noBreak"
          $ 1798 "movej(pose_trans(FRM_Reference, PSE_A), r=0.020)"
          movej( pose_trans (FRM_Reference, PSE_A), r=0.020)
        end
      end
      $ 1799 "MoveL"
      $ 1800 "If PSE_T_H≠PSE_Z"
      if (PSE_T_H != PSE_Z):
        $ 1801 "PSE_T_H" "breakAfter"
        movel(pose_trans(FRM_Reference, PSE_T_H), a=0.5, v=0.4, r=0.01)
      end
      $ 1802 "PSE_T" "breakAfter"
      global move_thread_flag_1802=0
      thread move_thread_1802():
        enter_critical
        move_thread_flag_1802 = 1
        movel(pose_trans(FRM_Reference, PSE_T), a=0.05, v=0.09)
        move_thread_flag_1802 = 2
        exit_critical
      end
      move_thread_flag_1802 = 0
      move_thread_han_1802 = run move_thread_1802()
      while (True):
        local targetTcpDirection=get_target_tcp_speed()
        local stepsToRetract=tool_contact(direction=targetTcpDirection)
        if (stepsToRetract > 0):
          kill move_thread_han_1802
          stopl(0.5)
          $ 1803 "Until (tool_contact_detection)"
          break
        end
        sleep(1.0E-10)
        if (move_thread_flag_1802 > 1):
          join move_thread_han_1802
          break
        end
        sync()
      end
      $ 1804 "Force"
      sleep(0.02)
      zero_ftsensor()
      force_mode(FRM_Reference, [1, 1, 1, 0, 0, 0], [0.0, 0.0, 0.0, 0.0, 0.0, 0.0], 2, [0.1, 0.1, 0.01, 0.3490658503988659, 0.3490658503988659, 0.3490658503988659])
      $ 1805 "PSE_T" "noBreak"
      movel(pose_trans(FRM_Reference, PSE_T), a=0.04, v=0.07)
      end_force_mode()
      stopl(5.0)
      $ 1806 "EXTT"
      $ 1807 "Switch JIG"
      switch_2 = JIG
      $ 1808 "Case 1"
      if (1 == switch_2):
        $ 1809 "3FG"
        $ 1810 "If OBJ_Picked"
        if (OBJ_Picked):
          $ 1811 "Set GRP_3F_Open=Off"
          set_standard_digital_out(5, False)
          $ 1812 "Wait: 0.2"
          sleep(0.2)
        end
      end
      $ 1813 "EOAT"
      $ 1814 "rq_move_and_wait_mm(GRP_Open_Pos)"
       rq_move_and_wait_mm (GRP_Open_Pos)
      $ 1815 "OBJ_Picked≔rq_is_object_detected()"
      global OBJ_Picked= rq_is_object_detected ()
      $ 1816 "If PSE_R_H≠PSE_Z"
      if (PSE_R_H != PSE_Z):
        $ 1817 "PSE_R" "breakAfter"
        movel(pose_trans(FRM_Reference, PSE_R), a=0.5, v=0.4, r=0.01)
        $ 1818 "PSE_R_H" "breakAfter"
        movel(pose_trans(FRM_Reference, PSE_R_H), a=0.5, v=0.4)
      else:
        $ 1819 "Else" "noBreak"
        $ 1820 "PSE_R" "breakAfter"
        movel(pose_trans(FRM_Reference, PSE_R), a=0.5, v=0.4)
      end
    elif (3 == switch_1):
      $ 1821 "Case 3"
      $ 1822 "Push"
      $ 1823 "Action_Info≔'push'"
      global Action_Info="push"
    elif (4 == switch_1):
      $ 1824 "Case 4"
      $ 1825 "Pull"
      $ 1826 "Action_Info≔'pull'"
      global Action_Info="pull"
    elif (6 == switch_1):
      $ 1829 "Case 6"
      $ 1830 "Drop the cap"
      $ 1831 "If JNT_A≠[0,0,0,0,0,0]"
      if (JNT_A != [0,0,0,0,0,0]):
        $ 1832 "MoveJ"
        $ 1833 "JNT_A" "breakAfter"
        movej(JNT_A, a=1.3962634015954636, v=1.7453292519943295, r=0.02)
      else:
        $ 1834 "Else" "noBreak"
        $ 1835 "MoveJ"
        $ 1836 "PSE_A" "breakAfter"
        movej(pose_trans(FRM_Reference, PSE_A), a=1.3962634015954636, v=1.7453292519943295, r=0.02)
      end
      $ 1837 "MoveL"
      $ 1838 "PSE_T" "breakAfter"
      movel(pose_trans(FRM_Reference, PSE_T), a=0.05, v=0.09)
      $ 1839 "'ADD OPEN GRIPPER'"
      # 'ADD OPEN GRIPPER'
      # begin: URCap Program Node
      #   Source: Robotiq_Grippers, 3.17.0.105337, Robotiq Inc.
      #   Type: Gripper
      $ 1840 "Gripper Move10mm (1)"
      if not(gripper_connected[0]):
        popup("Gripper 1 must be connected to run this program.", "No connection", False, True, True)
      end
      if not(rq_is_gripper_activated("1")):
        popup("Gripper 1 is not activated. Go to Installation tab > Gripper to activate it and run the program again.", "Not activated", False, True, True)
      end
      rq_set_pos_spd_for(201, 0, 28, "1")
      rq_wait_pos_spe_for_request(201, 0, 28, "1")
      rq_go_to("1")
      rq_wait("1")
      # end: URCap Program Node
      $ 1841 "PSE_T_H" "breakAfter"
      movel(pose_trans(FRM_Reference, PSE_T_H), a=0.05, v=0.09)
      # begin: URCap Program Node
      #   Source: Robotiq_Grippers, 3.17.0.105337, Robotiq Inc.
      #   Type: Gripper
      $ 1842 "Gripper Move40mm (1)"
      if not(gripper_connected[0]):
        popup("Gripper 1 must be connected to run this program.", "No connection", False, True, True)
      end
      if not(rq_is_gripper_activated("1")):
        popup("Gripper 1 is not activated. Go to Installation tab > Gripper to activate it and run the program again.", "Not activated", False, True, True)
      end
      rq_set_pos_spd_for(63, 0, 28, "1")
      rq_wait_pos_spe_for_request(63, 0, 28, "1")
      rq_go_to("1")
      rq_wait("1")
      # end: URCap Program Node
      $ 1843 "PSE_R" "breakAfter"
      movel(pose_trans(FRM_Reference, PSE_R), a=0.5, v=0.4)
    elif (7 == switch_1):
      $ 1844 "Case 7"
      $ 1845 "Load"
      $ 1846 "Action_Info≔'load object'"
      global Action_Info="load object"
      $ 1847 "do_transition(pose_trans(FRM_Reference, PSE_T), keep_rxry=OBJ_Picked)"
      do_transition( pose_trans (FRM_Reference, PSE_T), keep_rxry=OBJ_Picked)
      $ 1848 "If PSE_A_H≠PSE_Z"
      if (PSE_A_H != PSE_Z):
        $ 1849 "If JNT_Q≠JNT_Z"
        if (JNT_Q != JNT_Z):
          $ 1850 "movej(get_inverse_kin(pose_trans(FRM_Reference, PSE_A_H), qnear=JNT_Q), r=0.050)"
          movej(get_inverse_kin( pose_trans (FRM_Reference, PSE_A_H), qnear=JNT_Q), r=0.050)
        else:
          $ 1851 "Else" "noBreak"
          $ 1852 "movej(pose_trans(FRM_Reference, PSE_A_H), r=0.050)"
          movej( pose_trans (FRM_Reference, PSE_A_H), r=0.050)
        end
      end
      $ 1853 "If PSE_A≠PSE_Z"
      if (PSE_A != PSE_Z):
        $ 1854 "If JNT_Q≠JNT_Z"
        if (JNT_Q != JNT_Z):
          $ 1855 "movej(get_inverse_kin(pose_trans(FRM_Reference, PSE_A), qnear=JNT_Q), r=0.020)"
          movej(get_inverse_kin( pose_trans (FRM_Reference, PSE_A), qnear=JNT_Q), r=0.020)
        else:
          $ 1856 "Else" "noBreak"
          $ 1857 "movej(pose_trans(FRM_Reference, PSE_A), r=0.020)"
          movej( pose_trans (FRM_Reference, PSE_A), r=0.020)
        end
      end
      $ 1858 "MoveL"
      $ 1859 "If PSE_T_H≠PSE_Z"
      if (PSE_T_H != PSE_Z):
        $ 1860 "PSE_T_H" "breakAfter"
        movel(pose_trans(FRM_Reference, PSE_T_H), a=0.5, v=0.4, r=0.01)
      end
      $ 1861 "PSE_T" "breakAfter"
      global move_thread_flag_1861=0
      thread move_thread_1861():
        enter_critical
        move_thread_flag_1861 = 1
        movel(pose_trans(FRM_Reference, PSE_T), a=0.05, v=0.09)
        move_thread_flag_1861 = 2
        exit_critical
      end
      move_thread_flag_1861 = 0
      move_thread_han_1861 = run move_thread_1861()
      while (True):
        local targetTcpDirection=get_target_tcp_speed()
        local stepsToRetract=tool_contact(direction=targetTcpDirection)
        if (stepsToRetract > 0):
          kill move_thread_han_1861
          stopl(0.5)
          $ 1862 "Until (tool_contact_detection)"
          break
        end
        sleep(1.0E-10)
        if (move_thread_flag_1861 > 1):
          join move_thread_han_1861
          break
        end
        sync()
      end
      $ 1863 "Force"
      sleep(0.02)
      zero_ftsensor()
      force_mode(FRM_Reference, [0, 1, 1, 0, 0, 1], [0.0, 0.0, 0.0, 0.0, 0.0, 0.0], 2, [0.1, 0.05, 0.02, 0.3490658503988659, 0.3490658503988659, 3.141592653589793])
      $ 1864 "PSE_T" "noBreak"
      movel(pose_trans(FRM_Reference, PSE_T), a=0.04, v=0.07)
      end_force_mode()
      stopl(5.0)
      $ 1865 "EOAT"
      $ 1866 "rq_move_and_wait_mm(GRP_Open_Pos)"
       rq_move_and_wait_mm (GRP_Open_Pos)
      $ 1867 "OBJ_Picked≔rq_is_object_detected()"
      global OBJ_Picked= rq_is_object_detected ()
      $ 1868 "If PSE_R_H≠PSE_Z"
      if (PSE_R_H != PSE_Z):
        $ 1869 "PSE_R" "breakAfter"
        movel(pose_trans(FRM_Reference, PSE_R), a=0.5, v=0.4, r=0.01)
        $ 1870 "PSE_R_H" "breakAfter"
        movel(pose_trans(FRM_Reference, PSE_R_H), a=0.5, v=0.4)
      else:
        $ 1871 "Else" "noBreak"
        $ 1872 "PSE_R" "breakAfter"
        movel(pose_trans(FRM_Reference, PSE_R), a=0.5, v=0.4)
      end
    elif (8 == switch_1):
      $ 1873 "Case 8"
      $ 1874 "Unload"
      $ 1875 "Action_Info≔'pick object'"
      global Action_Info="pick object"
      $ 1876 "do_transition(pose_trans(FRM_Reference, PSE_T), keep_rxry=OBJ_Picked)"
      do_transition( pose_trans (FRM_Reference, PSE_T), keep_rxry=OBJ_Picked)
      $ 1877 "EOAT"
      $ 1878 "If  not OBJ_Picked"
      if (  not  OBJ_Picked):
        $ 1879 "rq_move_and_wait_mm(GRP_Open_Pos)"
         rq_move_and_wait_mm (GRP_Open_Pos)
      end
      $ 1880 "If PSE_A_H≠PSE_Z"
      if (PSE_A_H != PSE_Z):
        $ 1881 "If JNT_Q≠JNT_Z"
        if (JNT_Q != JNT_Z):
          $ 1882 "movej(get_inverse_kin(pose_trans(FRM_Reference, PSE_A_H), qnear=JNT_Q), r=0.050)"
          movej(get_inverse_kin( pose_trans (FRM_Reference, PSE_A_H), qnear=JNT_Q), r=0.050)
        else:
          $ 1883 "Else" "noBreak"
          $ 1884 "movej(pose_trans(FRM_Reference, PSE_A_H), r=0.050)"
          movej( pose_trans (FRM_Reference, PSE_A_H), r=0.050)
        end
      end
      $ 1885 "If PSE_A≠PSE_Z"
      if (PSE_A != PSE_Z):
        $ 1886 "If JNT_Q≠JNT_Z"
        if (JNT_Q != JNT_Z):
          $ 1887 "movej(get_inverse_kin(pose_trans(FRM_Reference, PSE_A), qnear=JNT_Q), r=0.020)"
          movej(get_inverse_kin( pose_trans (FRM_Reference, PSE_A), qnear=JNT_Q), r=0.020)
        else:
          $ 1888 "Else" "noBreak"
          $ 1889 "movej(pose_trans(FRM_Reference, PSE_A), r=0.020)"
          movej( pose_trans (FRM_Reference, PSE_A), r=0.020)
        end
      end
      $ 1890 "MoveL"
      $ 1891 "If PSE_T_H≠PSE_Z"
      if (PSE_T_H != PSE_Z):
        $ 1892 "PSE_T_H" "breakAfter"
        movel(pose_trans(FRM_Reference, PSE_T_H), a=0.5, v=0.4, r=0.01)
      end
      $ 1893 "PSE_T" "breakAfter"
      movel(pose_trans(FRM_Reference, PSE_T), a=0.08, v=0.12)
      $ 1894 "Force"
      sleep(0.02)
      zero_ftsensor()
      force_mode(FRM_Reference, [1, 1, 0, 0, 0, 0], [0.0, 0.0, 0.0, 0.0, 0.0, 0.0], 2, [0.05, 0.05, 0.1, 0.3490658503988659, 0.3490658503988659, 0.3490658503988659])
      $ 1895 "EOAT" "noBreak"
      $ 1896 "rq_set_force_norm(50)" "noBreak"
       rq_set_force_norm (50)
      $ 1897 "rq_close_and_wait()" "noBreak"
       rq_close_and_wait ()
      $ 1898 "OBJ_Picked≔rq_is_object_detected()" "noBreak"
      global OBJ_Picked= rq_is_object_detected ()
      $ 1899 "If  not OBJ_Picked" "noBreak"
      if (  not  OBJ_Picked):
        $ 1900 "set_error(ERROR_NO_OBJECT_TO_PICK)" "noBreak"
        set_error(ERROR_NO_OBJECT_TO_PICK)
      end
      $ 1901 "If PSE_R_H≠PSE_Z" "noBreak"
      if (PSE_R_H != PSE_Z):
        $ 1902 "PSE_R" "noBreak"
        movel(pose_trans(FRM_Reference, PSE_R), a=0.5, v=0.4, r=0.01)
        $ 1903 "PSE_R_H" "noBreak"
        movel(pose_trans(FRM_Reference, PSE_R_H), a=0.5, v=0.4)
      else:
        $ 1904 "Else" "noBreak"
        $ 1905 "PSE_R" "noBreak"
        movel(pose_trans(FRM_Reference, PSE_R), a=0.5, v=0.4)
      end
      end_force_mode()
      stopl(5.0)
    elif (11 == switch_1):
      $ 1906 "Case 11"
    elif (12 == switch_1):
      $ 1943 "Case 12"
      $ 1944 "Decap"
      $ 1945 "Action_Info≔'decapping'"
      global Action_Info="decapping"
      $ 1946 "Set GRP_3F_Enable=On"
      set_standard_digital_out(4, True)
      $ 1947 "Set GRP_3F_Decap=On"
      set_standard_digital_out(3, True)
      $ 1948 "Force"
      sleep(0.02)
      zero_ftsensor()
      force_mode(tool_pose(), [0, 0, 1, 0, 0, 0], [0.0, 0.0, 5.0, 0.0, 0.0, 0.0], 2, [0.1, 0.1, 0.15, 0.3490658503988659, 0.3490658503988659, 0.3490658503988659])
      $ 1949 "check_decapping(offset=0.015, timeout=5, abort=CMD_Hold)" "noBreak"
      check_decapping(offset=0.015, timeout=5, abort=CMD_Hold)
      end_force_mode()
      stopl(5.0)
      $ 1950 "Set GRP_3F_Decap=Off"
      set_standard_digital_out(3, False)
      $ 1951 "Set GRP_3F_Enable=Off"
      set_standard_digital_out(4, False)
      $ 1952 "MoveL"
      $ 1953 "PSE_R" "breakAfter"
      movel(pose_trans(FRM_Reference, PSE_R), a=0.8, v=0.15)
    elif (13 == switch_1):
      $ 1954 "Case 13"
      $ 1955 "TMR_Barcode: Reset"
      TMR_Barcode = 0
      $ 1956 "Read"
      $ 1957 "TMR_Barcode: Start"
      TMR_Barcode_is_counting = True
      $ 1958 "If TMR_Barcode<PRM_TO_Read_BC"
      global thread_flag_1958=0
      thread Thread_if_1958():
        $ 1959 "KeyenceTrigger"
        $ 1960 "Set OClearResult=HI:Pulse 0.2"
        thread SinglePulse14():
          write_output_boolean_register(2, True)
          sleep(0.2)
          write_output_boolean_register(2, False)
        end
        singlePulse14 = run SinglePulse14()
        $ 1961 "Wait: 0.5"
        sleep(0.5)
        $ 1962 "Set OTriggerBarcode=Off"
        write_output_boolean_register(1, False)
        $ 1963 "Wait: 0.5"
        sleep(0.5)
        $ 1964 "Set OTriggerBarcode=On"
        write_output_boolean_register(1, True)
        $ 1965 "Wait: 0.5"
        sleep(0.5)
        $ 1966 "Preorient"
        $ 1967 "TMR_Barcode: Reset"
        TMR_Barcode = 0
        $ 1968 "If ICmdExctd"
        if (read_input_boolean_register(12)):
          $ 1969 "Set GRP_3F_Decap=On"
          set_standard_digital_out(3, True)
          $ 1970 "Set GRP_3F_Enable=On"
          set_standard_digital_out(4, True)
          $ 1971 "Loop ICmdExctd"
          while (read_input_boolean_register(12)):
            $ 1972 "KeyenceTrigger"
            $ 1973 "Set OClearResult=HI:Pulse 0.1"
            thread SinglePulse15():
              write_output_boolean_register(2, True)
              sleep(0.1)
              write_output_boolean_register(2, False)
            end
            singlePulse15 = run SinglePulse15()
            $ 1974 "Wait: 0.3"
            sleep(0.3)
            $ 1975 "Set OTriggerBarcode=Off"
            write_output_boolean_register(1, False)
            $ 1976 "Wait: 0.3"
            sleep(0.3)
            $ 1977 "Set OTriggerBarcode=On"
            write_output_boolean_register(1, True)
            $ 1978 "Wait: 0.1"
            sleep(0.1)
          end
        end
        $ 1979 "If  not ICmdExctd"
        if (  not  read_input_boolean_register(12)):
          $ 1980 "Set GRP_3F_Decap=On"
          set_standard_digital_out(3, True)
          $ 1981 "Set GRP_3F_Enable=On"
          set_standard_digital_out(4, True)
          $ 1982 "Wait ICmdExctd=HI"
          while (read_input_boolean_register(12) == False):
            sync()
          end
        end
        $ 1983 "Set GRP_3F_Decap=Off"
        set_standard_digital_out(3, False)
        $ 1984 "Set GRP_3F_Enable=Off"
        set_standard_digital_out(4, False)
        $ 1985 "OBJ_Brc_OK≔ True "
        global OBJ_Brc_OK=  True
        thread_flag_1958 = 1
      end
      if (TMR_Barcode<PRM_TO_Read_BC):
        global thread_handler_1958=run Thread_if_1958()
        while (thread_flag_1958 == 0):
          if not(TMR_Barcode<PRM_TO_Read_BC):
            kill thread_handler_1958
            thread_flag_1958 = 2
          else:
            sync()
          end
        end
      else:
        thread_flag_1958 = 2
      end
      if (thread_flag_1958 == 2):
        $ 1986 "Else" "noBreak"
        $ 1987 "exeption"
        $ 1988 "error"
        $ 1990 "OBJ_Brc_OK≔ False "
        global OBJ_Brc_OK=  False
      end
      $ 1991 "Set GRP_3F_Decap=Off"
      set_standard_digital_out(3, False)
      $ 1992 "Set GRP_3F_Enable=Off"
      set_standard_digital_out(4, False)
      $ 1993 "Set OTriggerBarcode=Off"
      write_output_boolean_register(1, False)
    elif (15 == switch_1):
      $ 1994 "Case 15"
      $ 1995 "Detect"
      $ 1996 "Action_Info≔'detect'"
      global Action_Info="detect"
    elif (30 == switch_1):
      $ 1997 "Case 30"
      $ 1998 "Shake"
      $ 1999 "Action_Info≔'shake'"
      global Action_Info="shake"
      $ 2000 "do_transition(pose_trans(FRM_Reference, PSE_T), keep_rxry=OBJ_Picked)"
      do_transition( pose_trans (FRM_Reference, PSE_T), keep_rxry=OBJ_Picked)
      $ 2001 "If PSE_A_H≠PSE_Z"
      if (PSE_A_H != PSE_Z):
        $ 2002 "If JNT_Q≠JNT_Z"
        if (JNT_Q != JNT_Z):
          $ 2003 "movej(get_inverse_kin(pose_trans(FRM_Reference, PSE_A_H), qnear=JNT_Q), r=0.050)"
          movej(get_inverse_kin( pose_trans (FRM_Reference, PSE_A_H), qnear=JNT_Q), r=0.050)
        else:
          $ 2004 "Else" "noBreak"
          $ 2005 "movej(pose_trans(FRM_Reference, PSE_A_H), r=0.050)"
          movej( pose_trans (FRM_Reference, PSE_A_H), r=0.050)
        end
      end
      $ 2006 "If PSE_A≠PSE_Z"
      if (PSE_A != PSE_Z):
        $ 2007 "If JNT_Q≠JNT_Z"
        if (JNT_Q != JNT_Z):
          $ 2008 "movej(get_inverse_kin(pose_trans(FRM_Reference, PSE_A), qnear=JNT_Q), r=0.020)"
          movej(get_inverse_kin( pose_trans (FRM_Reference, PSE_A), qnear=JNT_Q), r=0.020)
        else:
          $ 2009 "Else" "noBreak"
          $ 2010 "movej(pose_trans(FRM_Reference, PSE_A), r=0.020)"
          movej( pose_trans (FRM_Reference, PSE_A), r=0.020)
        end
      end
      $ 2011 "MoveL"
      $ 2012 "If PSE_T_H≠PSE_Z"
      if (PSE_T_H != PSE_Z):
        $ 2013 "PSE_T_H" "breakAfter"
        movel(pose_trans(FRM_Reference, PSE_T_H), a=0.5, v=0.4, r=0.01)
      end
      $ 2014 "PSE_T" "breakAfter"
      movel(pose_trans(FRM_Reference, PSE_T), a=0.08, v=0.12)
      $ 2015 "EXTT"
      $ 2016 "Comment"
      # Comment
      $ 2017 "MoveJ"
      $ 2018 "Waypoint_54" "breakAfter"
      movej(get_inverse_kin(Waypoint_54_p, qnear=Waypoint_54_q), a=1.3962634015954636, v=1.0471975511965976)
      $ 2019 "MoveJ"
      $ 2020 "Waypoint_77" "breakAfter"
      movej(get_inverse_kin(Waypoint_77_p, qnear=Waypoint_77_q), a=1.3962634015954636, v=1.0471975511965976)
      $ 2021 "MoveJ"
      $ 2022 "Waypoint_83" "breakAfter"
      movej(get_inverse_kin(Waypoint_83_p, qnear=Waypoint_83_q), a=1.3962634015954636, v=1.0471975511965976)
      $ 2023 "MoveJ"
      $ 2024 "Waypoint_84" "breakAfter"
      movej(get_inverse_kin(Waypoint_84_p, qnear=Waypoint_84_q), a=1.3962634015954636, v=1.0471975511965976)
      $ 2025 "If PSE_R_H≠PSE_Z"
      if (PSE_R_H != PSE_Z):
        $ 2026 "PSE_R" "breakAfter"
        movel(pose_trans(FRM_Reference, PSE_R), a=0.5, v=0.4, r=0.01)
        $ 2027 "PSE_R_H" "breakAfter"
        movel(pose_trans(FRM_Reference, PSE_R_H), a=0.5, v=0.4)
      else:
        $ 2028 "Else" "noBreak"
        $ 2029 "PSE_R" "breakAfter"
        movel(pose_trans(FRM_Reference, PSE_R), a=0.5, v=0.4)
      end
    elif (31 == switch_1):
      $ 2030 "Case 31"
      $ 2031 "Action_Info≔'Pick_Vial'"
      global Action_Info="Pick_Vial"
      $ 2032 "Pick_Vial"
      # begin: URCap Program Node
      #   Source: Robotiq_Grippers, 3.17.0.105337, Robotiq Inc.
      #   Type: Gripper
      $ 2033 "Gripper Open (1)"
      if not(gripper_connected[0]):
        popup("Gripper 1 must be connected to run this program.", "No connection", False, True, True)
      end
      if not(rq_is_gripper_activated("1")):
        popup("Gripper 1 is not activated. Go to Installation tab > Gripper to activate it and run the program again.", "Not activated", False, True, True)
      end
      rq_set_pos_spd_for(0, 82, 71, "1")
      rq_wait_pos_spe_for_request(0, 82, 71, "1")
      rq_go_to("1")
      rq_wait("1")
      # end: URCap Program Node
      $ 2034 "MoveJ"
      $ 2035 "Vial_above_1" "breakAfter"
      movej(get_inverse_kin(Vial_above_1_p, qnear=Vial_above_1_q), a=0.5235987755982988, v=0.4363323129985824, r=0.05)
      $ 2036 "MoveL"
      $ 2037 "Vial_pick_poi_1" "breakAfter"
      movel(Vial_pick_poi_1_p, a=0.5, v=0.1)
      # begin: URCap Program Node
      #   Source: Robotiq_Grippers, 3.17.0.105337, Robotiq Inc.
      #   Type: Gripper
      $ 2038 "Gripper Close (1)"
      if not(gripper_connected[0]):
        popup("Gripper 1 must be connected to run this program.", "No connection", False, True, True)
      end
      if not(rq_is_gripper_activated("1")):
        popup("Gripper 1 is not activated. Go to Installation tab > Gripper to activate it and run the program again.", "Not activated", False, True, True)
      end
      rq_set_pos_spd_for(255, 71, 84, "1")
      rq_wait_pos_spe_for_request(255, 71, 84, "1")
      rq_go_to("1")
      rq_wait("1")
      # end: URCap Program Node
      $ 2039 "MoveL"
      $ 2040 "Waypoint_86" "breakAfter"
      movel(Waypoint_86_p, a=0.5, v=0.1, r=0.05)
      $ 2041 "Home (Safe)"
      movej([-1.2302089344500047, -1.2969853503591224, -1.875639182904262, -1.539621866126728, 1.5731943360401213, -2.80099559440227], a=1.3962634015954636, v=1.0471975511965976)
    elif (32 == switch_1):
      $ 2042 "Case 32"
      $ 2044 "decap_Vial"
      $ 2045 "Set GRP_3F_Open=On"
      set_standard_digital_out(5, True)
      $ 2046 "MoveJ"
      $ 2047 "Waypoint_87" "breakAfter"
      movej(get_inverse_kin(Waypoint_87_p, qnear=Waypoint_87_q), a=0.5235987755982988, v=0.4363323129985824)
      $ 2048 "MoveL"
      $ 2049 "Vial_3FG_plac_1" "breakAfter"
      movel(Vial_3FG_plac_1_p, a=0.5, v=0.1)
      $ 2050 "Set GRP_3F_Open=Off"
